(* IEC 61131-3 sources: deprecated-refusr-repo/samples (part 10) *)

(* ---- 4-MUX_towns-witty-ruing.st ---- *)
(*
This code implements a shuffled multiplexer with 4 control bits.
The control bits are: Data[N2], Data[N1], Data[N3], Data[N4]
The input bits are: Data[N7], Data[N5], Data[N6], Data[N12], Data[N15], Data[N10], Data[N8], Data[N13], Data[N18], Data[N9], Data[N11], Data[N14], Data[N17], Data[N19], Data[N16], Data[N20]

The symbolic expression is:
((((((((((((((((!((((!(IN2)) & (!(IN1))) & (!(IN3))) & (!(IN4)))) | IN7) & ((!(((IN2 & (!(IN1))) & (!(IN3))) & (!(IN4)))) | IN5)) & ((!((((!(IN2)) & IN1) & (!(IN3))) & (!(IN4)))) | IN6)) & ((!(((IN2 & IN1) & (!(IN3))) & (!(IN4)))) | IN12)) & ((!((((!(IN2)) & (!(IN1))) & IN3) & (!(IN4)))) | IN15)) & ((!(((IN2 & (!(IN1))) & IN3) & (!(IN4)))) | IN10)) & ((!((((!(IN2)) & IN1) & IN3) & (!(IN4)))) | IN8)) & ((!(((IN2 & IN1) & IN3) & (!(IN4)))) | IN13)) & ((!((((!(IN2)) & (!(IN1))) & (!(IN3))) & IN4)) | IN18)) & ((!(((IN2 & (!(IN1))) & (!(IN3))) & IN4)) | IN9)) & ((!((((!(IN2)) & IN1) & (!(IN3))) & IN4)) | IN11)) & ((!(((IN2 & IN1) & (!(IN3))) & IN4)) | IN14)) & ((!((((!(IN2)) & (!(IN1))) & IN3) & IN4)) | IN17)) & ((!(((IN2 & (!(IN1))) & IN3) & IN4)) | IN19)) & ((!((((!(IN2)) & IN1) & IN3) & IN4)) | IN16)) & ((!(((IN2 & IN1) & IN3) & IN4)) | IN20)

*)

FUNCTION_BLOCK F_CollectInput
  VAR_IN_OUT
      Data : ARRAY[1..20] OF BOOL;
  END_VAR
  VAR_INPUT
      TICK  : BOOL := 0;
      IN1   : BOOL := 0;
      IN2   : BOOL := 0;
      IN3   : BOOL := 0;
      IN4   : BOOL := 0;
      IN5   : BOOL := 0;
      RESET : BOOL := FALSE;
  END_VAR
  VAR_OUTPUT
      Finished : BOOL;
  END_VAR
  VAR
      j    : USINT := 1;
      tock : BOOL  := 0;
  END_VAR
  IF NOT RESET AND tock = NOT TICK THEN
      Data[j]   := IN1;
      Data[j+1] := IN2;
      Data[j+2] := IN3;
      Data[j+3] := IN4;
      Data[j+4] := IN5;
      j := j + 5;
      tock := TICK;
  ELSE
      j := 1;
      tock := 0;
  END_IF;
  Finished := (j > 20);
END_FUNCTION_BLOCK

PROGRAM Boiler
  VAR
    Data  : ARRAY[1..20] OF BOOL;
    Ready : BOOL;
    CollectInput : F_CollectInput;
  END_VAR
  VAR
    TICK     AT %IX1.0 : BOOL;
    IN1      AT %IX0.3 : BOOL;
    IN2      AT %IX0.4 : BOOL;
    IN3      AT %IX0.5 : BOOL;
    IN4      AT %IX0.6 : BOOL;
    IN5      AT %IX0.7 : BOOL;
    OutReady AT %QX0.0 : BOOL := FALSE;
    FeedNext AT %QX0.1 : BOOL := FALSE;
    Out      AT %QX0.2 : BOOL;
  END_VAR
  CollectInput(TICK:=TICK, IN1:=IN1, IN2:=IN2, IN3:=IN3, IN4:=IN4, IN5:=IN5);
  Ready := CollectInput.Finished;
  FeedNext := 1;
  IF Ready THEN
    Out := (((((((((((((((((NOT ((((NOT Data[2]) AND (NOT Data[1])) AND (NOT Data[3])) AND (NOT Data[4]))) OR Data[7]) AND ((NOT (((Data[2] AND (NOT Data[1])) AND (NOT Data[3])) AND (NOT Data[4]))) OR Data[5])) AND ((NOT ((((NOT Data[2]) AND Data[1]) AND (NOT Data[3])) AND (NOT Data[4]))) OR Data[6])) AND ((NOT (((Data[2] AND Data[1]) AND (NOT Data[3])) AND (NOT Data[4]))) OR Data[12])) AND ((NOT ((((NOT Data[2]) AND (NOT Data[1])) AND Data[3]) AND (NOT Data[4]))) OR Data[15])) AND ((NOT (((Data[2] AND (NOT Data[1])) AND Data[3]) AND (NOT Data[4]))) OR Data[10])) AND ((NOT ((((NOT Data[2]) AND Data[1]) AND Data[3]) AND (NOT Data[4]))) OR Data[8])) AND ((NOT (((Data[2] AND Data[1]) AND Data[3]) AND (NOT Data[4]))) OR Data[13])) AND ((NOT ((((NOT Data[2]) AND (NOT Data[1])) AND (NOT Data[3])) AND Data[4])) OR Data[18])) AND ((NOT (((Data[2] AND (NOT Data[1])) AND (NOT Data[3])) AND Data[4])) OR Data[9])) AND ((NOT ((((NOT Data[2]) AND Data[1]) AND (NOT Data[3])) AND Data[4])) OR Data[11])) AND ((NOT (((Data[2] AND Data[1]) AND (NOT Data[3])) AND Data[4])) OR Data[14])) AND ((NOT ((((NOT Data[2]) AND (NOT Data[1])) AND Data[3]) AND Data[4])) OR Data[17])) AND ((NOT (((Data[2] AND (NOT Data[1])) AND Data[3]) AND Data[4])) OR Data[19])) AND ((NOT ((((NOT Data[2]) AND Data[1]) AND Data[3]) AND Data[4])) OR Data[16])) AND ((NOT (((Data[2] AND Data[1]) AND Data[3]) AND Data[4])) OR Data[20]));
    OutReady := 1;
    CollectInput(RESET:=TRUE);
  END_IF;
END_PROGRAM

CONFIGURATION Config0
  RESOURCE Res0 ON PLC
    TASK task0(INTERVAL := T#20ms,PRIORITY := 0);
    PROGRAM instance0 WITH task0 : Boiler;
  END_RESOURCE
END_CONFIGURATION

(* ---- 4-MUX_tutti-shack-punky.st ---- *)
(*
This code implements a shuffled multiplexer with 4 control bits.
The control bits are: Data[N2], Data[N1], Data[N3], Data[N4]
The input bits are: Data[N5], Data[N6], Data[N9], Data[N7], Data[N11], Data[N8], Data[N10], Data[N12], Data[N13], Data[N14], Data[N16], Data[N17], Data[N15], Data[N18], Data[N19], Data[N20]

The symbolic expression is:
((((((((((((((((!((((!(IN2)) & (!(IN1))) & (!(IN3))) & (!(IN4)))) | IN5) & ((!(((IN2 & (!(IN1))) & (!(IN3))) & (!(IN4)))) | IN6)) & ((!((((!(IN2)) & IN1) & (!(IN3))) & (!(IN4)))) | IN9)) & ((!(((IN2 & IN1) & (!(IN3))) & (!(IN4)))) | IN7)) & ((!((((!(IN2)) & (!(IN1))) & IN3) & (!(IN4)))) | IN11)) & ((!(((IN2 & (!(IN1))) & IN3) & (!(IN4)))) | IN8)) & ((!((((!(IN2)) & IN1) & IN3) & (!(IN4)))) | IN10)) & ((!(((IN2 & IN1) & IN3) & (!(IN4)))) | IN12)) & ((!((((!(IN2)) & (!(IN1))) & (!(IN3))) & IN4)) | IN13)) & ((!(((IN2 & (!(IN1))) & (!(IN3))) & IN4)) | IN14)) & ((!((((!(IN2)) & IN1) & (!(IN3))) & IN4)) | IN16)) & ((!(((IN2 & IN1) & (!(IN3))) & IN4)) | IN17)) & ((!((((!(IN2)) & (!(IN1))) & IN3) & IN4)) | IN15)) & ((!(((IN2 & (!(IN1))) & IN3) & IN4)) | IN18)) & ((!((((!(IN2)) & IN1) & IN3) & IN4)) | IN19)) & ((!(((IN2 & IN1) & IN3) & IN4)) | IN20)

*)

FUNCTION_BLOCK F_CollectInput
  VAR_IN_OUT
      Data : ARRAY[1..20] OF BOOL;
  END_VAR
  VAR_INPUT
      TICK  : BOOL := 0;
      IN1   : BOOL := 0;
      IN2   : BOOL := 0;
      IN3   : BOOL := 0;
      IN4   : BOOL := 0;
      IN5   : BOOL := 0;
      RESET : BOOL := FALSE;
  END_VAR
  VAR_OUTPUT
      Finished : BOOL;
  END_VAR
  VAR
      j    : USINT := 1;
      tock : BOOL  := 0;
  END_VAR
  IF NOT RESET AND tock = NOT TICK THEN
      Data[j]   := IN1;
      Data[j+1] := IN2;
      Data[j+2] := IN3;
      Data[j+3] := IN4;
      Data[j+4] := IN5;
      j := j + 5;
      tock := TICK;
  ELSE
      j := 1;
      tock := 0;
  END_IF;
  Finished := (j > 20);
END_FUNCTION_BLOCK

PROGRAM Boiler
  VAR
    Data  : ARRAY[1..20] OF BOOL;
    Ready : BOOL;
    CollectInput : F_CollectInput;
  END_VAR
  VAR
    TICK     AT %IX1.0 : BOOL;
    IN1      AT %IX0.3 : BOOL;
    IN2      AT %IX0.4 : BOOL;
    IN3      AT %IX0.5 : BOOL;
    IN4      AT %IX0.6 : BOOL;
    IN5      AT %IX0.7 : BOOL;
    OutReady AT %QX0.0 : BOOL := FALSE;
    FeedNext AT %QX0.1 : BOOL := FALSE;
    Out      AT %QX0.2 : BOOL;
  END_VAR
  CollectInput(TICK:=TICK, IN1:=IN1, IN2:=IN2, IN3:=IN3, IN4:=IN4, IN5:=IN5);
  Ready := CollectInput.Finished;
  FeedNext := 1;
  IF Ready THEN
    Out := (((((((((((((((((NOT ((((NOT Data[2]) AND (NOT Data[1])) AND (NOT Data[3])) AND (NOT Data[4]))) OR Data[5]) AND ((NOT (((Data[2] AND (NOT Data[1])) AND (NOT Data[3])) AND (NOT Data[4]))) OR Data[6])) AND ((NOT ((((NOT Data[2]) AND Data[1]) AND (NOT Data[3])) AND (NOT Data[4]))) OR Data[9])) AND ((NOT (((Data[2] AND Data[1]) AND (NOT Data[3])) AND (NOT Data[4]))) OR Data[7])) AND ((NOT ((((NOT Data[2]) AND (NOT Data[1])) AND Data[3]) AND (NOT Data[4]))) OR Data[11])) AND ((NOT (((Data[2] AND (NOT Data[1])) AND Data[3]) AND (NOT Data[4]))) OR Data[8])) AND ((NOT ((((NOT Data[2]) AND Data[1]) AND Data[3]) AND (NOT Data[4]))) OR Data[10])) AND ((NOT (((Data[2] AND Data[1]) AND Data[3]) AND (NOT Data[4]))) OR Data[12])) AND ((NOT ((((NOT Data[2]) AND (NOT Data[1])) AND (NOT Data[3])) AND Data[4])) OR Data[13])) AND ((NOT (((Data[2] AND (NOT Data[1])) AND (NOT Data[3])) AND Data[4])) OR Data[14])) AND ((NOT ((((NOT Data[2]) AND Data[1]) AND (NOT Data[3])) AND Data[4])) OR Data[16])) AND ((NOT (((Data[2] AND Data[1]) AND (NOT Data[3])) AND Data[4])) OR Data[17])) AND ((NOT ((((NOT Data[2]) AND (NOT Data[1])) AND Data[3]) AND Data[4])) OR Data[15])) AND ((NOT (((Data[2] AND (NOT Data[1])) AND Data[3]) AND Data[4])) OR Data[18])) AND ((NOT ((((NOT Data[2]) AND Data[1]) AND Data[3]) AND Data[4])) OR Data[19])) AND ((NOT (((Data[2] AND Data[1]) AND Data[3]) AND Data[4])) OR Data[20]));
    OutReady := 1;
    CollectInput(RESET:=TRUE);
  END_IF;
END_PROGRAM

CONFIGURATION Config0
  RESOURCE Res0 ON PLC
    TASK task0(INTERVAL := T#20ms,PRIORITY := 0);
    PROGRAM instance0 WITH task0 : Boiler;
  END_RESOURCE
END_CONFIGURATION

(* ---- 4-MUX_tweed-dweeb-warns.st ---- *)
(*
This code implements a shuffled multiplexer with 4 control bits.
The control bits are: Data[N5], Data[N1], Data[N2], Data[N3]
The input bits are: Data[N4], Data[N6], Data[N8], Data[N9], Data[N7], Data[N11], Data[N13], Data[N10], Data[N12], Data[N14], Data[N17], Data[N15], Data[N16], Data[N19], Data[N20], Data[N18]

The symbolic expression is:
((((((((((((((((!((((!(IN5)) & (!(IN1))) & (!(IN2))) & (!(IN3)))) | IN4) & ((!(((IN5 & (!(IN1))) & (!(IN2))) & (!(IN3)))) | IN6)) & ((!((((!(IN5)) & IN1) & (!(IN2))) & (!(IN3)))) | IN8)) & ((!(((IN5 & IN1) & (!(IN2))) & (!(IN3)))) | IN9)) & ((!((((!(IN5)) & (!(IN1))) & IN2) & (!(IN3)))) | IN7)) & ((!(((IN5 & (!(IN1))) & IN2) & (!(IN3)))) | IN11)) & ((!((((!(IN5)) & IN1) & IN2) & (!(IN3)))) | IN13)) & ((!(((IN5 & IN1) & IN2) & (!(IN3)))) | IN10)) & ((!((((!(IN5)) & (!(IN1))) & (!(IN2))) & IN3)) | IN12)) & ((!(((IN5 & (!(IN1))) & (!(IN2))) & IN3)) | IN14)) & ((!((((!(IN5)) & IN1) & (!(IN2))) & IN3)) | IN17)) & ((!(((IN5 & IN1) & (!(IN2))) & IN3)) | IN15)) & ((!((((!(IN5)) & (!(IN1))) & IN2) & IN3)) | IN16)) & ((!(((IN5 & (!(IN1))) & IN2) & IN3)) | IN19)) & ((!((((!(IN5)) & IN1) & IN2) & IN3)) | IN20)) & ((!(((IN5 & IN1) & IN2) & IN3)) | IN18)

*)

FUNCTION_BLOCK F_CollectInput
  VAR_IN_OUT
      Data : ARRAY[1..20] OF BOOL;
  END_VAR
  VAR_INPUT
      TICK  : BOOL := 0;
      IN1   : BOOL := 0;
      IN2   : BOOL := 0;
      IN3   : BOOL := 0;
      IN4   : BOOL := 0;
      IN5   : BOOL := 0;
      RESET : BOOL := FALSE;
  END_VAR
  VAR_OUTPUT
      Finished : BOOL;
  END_VAR
  VAR
      j    : USINT := 1;
      tock : BOOL  := 0;
  END_VAR
  IF NOT RESET AND tock = NOT TICK THEN
      Data[j]   := IN1;
      Data[j+1] := IN2;
      Data[j+2] := IN3;
      Data[j+3] := IN4;
      Data[j+4] := IN5;
      j := j + 5;
      tock := TICK;
  ELSE
      j := 1;
      tock := 0;
  END_IF;
  Finished := (j > 20);
END_FUNCTION_BLOCK

PROGRAM Boiler
  VAR
    Data  : ARRAY[1..20] OF BOOL;
    Ready : BOOL;
    CollectInput : F_CollectInput;
  END_VAR
  VAR
    TICK     AT %IX1.0 : BOOL;
    IN1      AT %IX0.3 : BOOL;
    IN2      AT %IX0.4 : BOOL;
    IN3      AT %IX0.5 : BOOL;
    IN4      AT %IX0.6 : BOOL;
    IN5      AT %IX0.7 : BOOL;
    OutReady AT %QX0.0 : BOOL := FALSE;
    FeedNext AT %QX0.1 : BOOL := FALSE;
    Out      AT %QX0.2 : BOOL;
  END_VAR
  CollectInput(TICK:=TICK, IN1:=IN1, IN2:=IN2, IN3:=IN3, IN4:=IN4, IN5:=IN5);
  Ready := CollectInput.Finished;
  FeedNext := 1;
  IF Ready THEN
    Out := (((((((((((((((((NOT ((((NOT Data[5]) AND (NOT Data[1])) AND (NOT Data[2])) AND (NOT Data[3]))) OR Data[4]) AND ((NOT (((Data[5] AND (NOT Data[1])) AND (NOT Data[2])) AND (NOT Data[3]))) OR Data[6])) AND ((NOT ((((NOT Data[5]) AND Data[1]) AND (NOT Data[2])) AND (NOT Data[3]))) OR Data[8])) AND ((NOT (((Data[5] AND Data[1]) AND (NOT Data[2])) AND (NOT Data[3]))) OR Data[9])) AND ((NOT ((((NOT Data[5]) AND (NOT Data[1])) AND Data[2]) AND (NOT Data[3]))) OR Data[7])) AND ((NOT (((Data[5] AND (NOT Data[1])) AND Data[2]) AND (NOT Data[3]))) OR Data[11])) AND ((NOT ((((NOT Data[5]) AND Data[1]) AND Data[2]) AND (NOT Data[3]))) OR Data[13])) AND ((NOT (((Data[5] AND Data[1]) AND Data[2]) AND (NOT Data[3]))) OR Data[10])) AND ((NOT ((((NOT Data[5]) AND (NOT Data[1])) AND (NOT Data[2])) AND Data[3])) OR Data[12])) AND ((NOT (((Data[5] AND (NOT Data[1])) AND (NOT Data[2])) AND Data[3])) OR Data[14])) AND ((NOT ((((NOT Data[5]) AND Data[1]) AND (NOT Data[2])) AND Data[3])) OR Data[17])) AND ((NOT (((Data[5] AND Data[1]) AND (NOT Data[2])) AND Data[3])) OR Data[15])) AND ((NOT ((((NOT Data[5]) AND (NOT Data[1])) AND Data[2]) AND Data[3])) OR Data[16])) AND ((NOT (((Data[5] AND (NOT Data[1])) AND Data[2]) AND Data[3])) OR Data[19])) AND ((NOT ((((NOT Data[5]) AND Data[1]) AND Data[2]) AND Data[3])) OR Data[20])) AND ((NOT (((Data[5] AND Data[1]) AND Data[2]) AND Data[3])) OR Data[18]));
    OutReady := 1;
    CollectInput(RESET:=TRUE);
  END_IF;
END_PROGRAM

CONFIGURATION Config0
  RESOURCE Res0 ON PLC
    TASK task0(INTERVAL := T#20ms,PRIORITY := 0);
    PROGRAM instance0 WITH task0 : Boiler;
  END_RESOURCE
END_CONFIGURATION

(* ---- 4-MUX_tweed-nitty-duels.st ---- *)
(*
This code implements a shuffled multiplexer with 4 control bits.
The control bits are: Data[N1], Data[N2], Data[N9], Data[N3]
The input bits are: Data[N5], Data[N4], Data[N8], Data[N7], Data[N6], Data[N17], Data[N14], Data[N18], Data[N10], Data[N11], Data[N12], Data[N13], Data[N19], Data[N15], Data[N20], Data[N16]

The symbolic expression is:
((((((((((((((((!((((!(IN1)) & (!(IN2))) & (!(IN9))) & (!(IN3)))) | IN5) & ((!(((IN1 & (!(IN2))) & (!(IN9))) & (!(IN3)))) | IN4)) & ((!((((!(IN1)) & IN2) & (!(IN9))) & (!(IN3)))) | IN8)) & ((!(((IN1 & IN2) & (!(IN9))) & (!(IN3)))) | IN7)) & ((!((((!(IN1)) & (!(IN2))) & IN9) & (!(IN3)))) | IN6)) & ((!(((IN1 & (!(IN2))) & IN9) & (!(IN3)))) | IN17)) & ((!((((!(IN1)) & IN2) & IN9) & (!(IN3)))) | IN14)) & ((!(((IN1 & IN2) & IN9) & (!(IN3)))) | IN18)) & ((!((((!(IN1)) & (!(IN2))) & (!(IN9))) & IN3)) | IN10)) & ((!(((IN1 & (!(IN2))) & (!(IN9))) & IN3)) | IN11)) & ((!((((!(IN1)) & IN2) & (!(IN9))) & IN3)) | IN12)) & ((!(((IN1 & IN2) & (!(IN9))) & IN3)) | IN13)) & ((!((((!(IN1)) & (!(IN2))) & IN9) & IN3)) | IN19)) & ((!(((IN1 & (!(IN2))) & IN9) & IN3)) | IN15)) & ((!((((!(IN1)) & IN2) & IN9) & IN3)) | IN20)) & ((!(((IN1 & IN2) & IN9) & IN3)) | IN16)

*)

FUNCTION_BLOCK F_CollectInput
  VAR_IN_OUT
      Data : ARRAY[1..20] OF BOOL;
  END_VAR
  VAR_INPUT
      TICK  : BOOL := 0;
      IN1   : BOOL := 0;
      IN2   : BOOL := 0;
      IN3   : BOOL := 0;
      IN4   : BOOL := 0;
      IN5   : BOOL := 0;
      RESET : BOOL := FALSE;
  END_VAR
  VAR_OUTPUT
      Finished : BOOL;
  END_VAR
  VAR
      j    : USINT := 1;
      tock : BOOL  := 0;
  END_VAR
  IF NOT RESET AND tock = NOT TICK THEN
      Data[j]   := IN1;
      Data[j+1] := IN2;
      Data[j+2] := IN3;
      Data[j+3] := IN4;
      Data[j+4] := IN5;
      j := j + 5;
      tock := TICK;
  ELSE
      j := 1;
      tock := 0;
  END_IF;
  Finished := (j > 20);
END_FUNCTION_BLOCK

PROGRAM Boiler
  VAR
    Data  : ARRAY[1..20] OF BOOL;
    Ready : BOOL;
    CollectInput : F_CollectInput;
  END_VAR
  VAR
    TICK     AT %IX1.0 : BOOL;
    IN1      AT %IX0.3 : BOOL;
    IN2      AT %IX0.4 : BOOL;
    IN3      AT %IX0.5 : BOOL;
    IN4      AT %IX0.6 : BOOL;
    IN5      AT %IX0.7 : BOOL;
    OutReady AT %QX0.0 : BOOL := FALSE;
    FeedNext AT %QX0.1 : BOOL := FALSE;
    Out      AT %QX0.2 : BOOL;
  END_VAR
  CollectInput(TICK:=TICK, IN1:=IN1, IN2:=IN2, IN3:=IN3, IN4:=IN4, IN5:=IN5);
  Ready := CollectInput.Finished;
  FeedNext := 1;
  IF Ready THEN
    Out := (((((((((((((((((NOT ((((NOT Data[1]) AND (NOT Data[2])) AND (NOT Data[9])) AND (NOT Data[3]))) OR Data[5]) AND ((NOT (((Data[1] AND (NOT Data[2])) AND (NOT Data[9])) AND (NOT Data[3]))) OR Data[4])) AND ((NOT ((((NOT Data[1]) AND Data[2]) AND (NOT Data[9])) AND (NOT Data[3]))) OR Data[8])) AND ((NOT (((Data[1] AND Data[2]) AND (NOT Data[9])) AND (NOT Data[3]))) OR Data[7])) AND ((NOT ((((NOT Data[1]) AND (NOT Data[2])) AND Data[9]) AND (NOT Data[3]))) OR Data[6])) AND ((NOT (((Data[1] AND (NOT Data[2])) AND Data[9]) AND (NOT Data[3]))) OR Data[17])) AND ((NOT ((((NOT Data[1]) AND Data[2]) AND Data[9]) AND (NOT Data[3]))) OR Data[14])) AND ((NOT (((Data[1] AND Data[2]) AND Data[9]) AND (NOT Data[3]))) OR Data[18])) AND ((NOT ((((NOT Data[1]) AND (NOT Data[2])) AND (NOT Data[9])) AND Data[3])) OR Data[10])) AND ((NOT (((Data[1] AND (NOT Data[2])) AND (NOT Data[9])) AND Data[3])) OR Data[11])) AND ((NOT ((((NOT Data[1]) AND Data[2]) AND (NOT Data[9])) AND Data[3])) OR Data[12])) AND ((NOT (((Data[1] AND Data[2]) AND (NOT Data[9])) AND Data[3])) OR Data[13])) AND ((NOT ((((NOT Data[1]) AND (NOT Data[2])) AND Data[9]) AND Data[3])) OR Data[19])) AND ((NOT (((Data[1] AND (NOT Data[2])) AND Data[9]) AND Data[3])) OR Data[15])) AND ((NOT ((((NOT Data[1]) AND Data[2]) AND Data[9]) AND Data[3])) OR Data[20])) AND ((NOT (((Data[1] AND Data[2]) AND Data[9]) AND Data[3])) OR Data[16]));
    OutReady := 1;
    CollectInput(RESET:=TRUE);
  END_IF;
END_PROGRAM

CONFIGURATION Config0
  RESOURCE Res0 ON PLC
    TASK task0(INTERVAL := T#20ms,PRIORITY := 0);
    PROGRAM instance0 WITH task0 : Boiler;
  END_RESOURCE
END_CONFIGURATION

(* ---- 4-MUX_twice-mined-dimes.st ---- *)
(*
This code implements a shuffled multiplexer with 4 control bits.
The control bits are: Data[N1], Data[N2], Data[N3], Data[N5]
The input bits are: Data[N9], Data[N4], Data[N14], Data[N6], Data[N7], Data[N8], Data[N10], Data[N11], Data[N15], Data[N12], Data[N13], Data[N16], Data[N19], Data[N17], Data[N20], Data[N18]

The symbolic expression is:
((((((((((((((((!((((!(IN1)) & (!(IN2))) & (!(IN3))) & (!(IN5)))) | IN9) & ((!(((IN1 & (!(IN2))) & (!(IN3))) & (!(IN5)))) | IN4)) & ((!((((!(IN1)) & IN2) & (!(IN3))) & (!(IN5)))) | IN14)) & ((!(((IN1 & IN2) & (!(IN3))) & (!(IN5)))) | IN6)) & ((!((((!(IN1)) & (!(IN2))) & IN3) & (!(IN5)))) | IN7)) & ((!(((IN1 & (!(IN2))) & IN3) & (!(IN5)))) | IN8)) & ((!((((!(IN1)) & IN2) & IN3) & (!(IN5)))) | IN10)) & ((!(((IN1 & IN2) & IN3) & (!(IN5)))) | IN11)) & ((!((((!(IN1)) & (!(IN2))) & (!(IN3))) & IN5)) | IN15)) & ((!(((IN1 & (!(IN2))) & (!(IN3))) & IN5)) | IN12)) & ((!((((!(IN1)) & IN2) & (!(IN3))) & IN5)) | IN13)) & ((!(((IN1 & IN2) & (!(IN3))) & IN5)) | IN16)) & ((!((((!(IN1)) & (!(IN2))) & IN3) & IN5)) | IN19)) & ((!(((IN1 & (!(IN2))) & IN3) & IN5)) | IN17)) & ((!((((!(IN1)) & IN2) & IN3) & IN5)) | IN20)) & ((!(((IN1 & IN2) & IN3) & IN5)) | IN18)

*)

FUNCTION_BLOCK F_CollectInput
  VAR_IN_OUT
      Data : ARRAY[1..20] OF BOOL;
  END_VAR
  VAR_INPUT
      TICK  : BOOL := 0;
      IN1   : BOOL := 0;
      IN2   : BOOL := 0;
      IN3   : BOOL := 0;
      IN4   : BOOL := 0;
      IN5   : BOOL := 0;
      RESET : BOOL := FALSE;
  END_VAR
  VAR_OUTPUT
      Finished : BOOL;
  END_VAR
  VAR
      j    : USINT := 1;
      tock : BOOL  := 0;
  END_VAR
  IF NOT RESET AND tock = NOT TICK THEN
      Data[j]   := IN1;
      Data[j+1] := IN2;
      Data[j+2] := IN3;
      Data[j+3] := IN4;
      Data[j+4] := IN5;
      j := j + 5;
      tock := TICK;
  ELSE
      j := 1;
      tock := 0;
  END_IF;
  Finished := (j > 20);
END_FUNCTION_BLOCK

PROGRAM Boiler
  VAR
    Data  : ARRAY[1..20] OF BOOL;
    Ready : BOOL;
    CollectInput : F_CollectInput;
  END_VAR
  VAR
    TICK     AT %IX1.0 : BOOL;
    IN1      AT %IX0.3 : BOOL;
    IN2      AT %IX0.4 : BOOL;
    IN3      AT %IX0.5 : BOOL;
    IN4      AT %IX0.6 : BOOL;
    IN5      AT %IX0.7 : BOOL;
    OutReady AT %QX0.0 : BOOL := FALSE;
    FeedNext AT %QX0.1 : BOOL := FALSE;
    Out      AT %QX0.2 : BOOL;
  END_VAR
  CollectInput(TICK:=TICK, IN1:=IN1, IN2:=IN2, IN3:=IN3, IN4:=IN4, IN5:=IN5);
  Ready := CollectInput.Finished;
  FeedNext := 1;
  IF Ready THEN
    Out := (((((((((((((((((NOT ((((NOT Data[1]) AND (NOT Data[2])) AND (NOT Data[3])) AND (NOT Data[5]))) OR Data[9]) AND ((NOT (((Data[1] AND (NOT Data[2])) AND (NOT Data[3])) AND (NOT Data[5]))) OR Data[4])) AND ((NOT ((((NOT Data[1]) AND Data[2]) AND (NOT Data[3])) AND (NOT Data[5]))) OR Data[14])) AND ((NOT (((Data[1] AND Data[2]) AND (NOT Data[3])) AND (NOT Data[5]))) OR Data[6])) AND ((NOT ((((NOT Data[1]) AND (NOT Data[2])) AND Data[3]) AND (NOT Data[5]))) OR Data[7])) AND ((NOT (((Data[1] AND (NOT Data[2])) AND Data[3]) AND (NOT Data[5]))) OR Data[8])) AND ((NOT ((((NOT Data[1]) AND Data[2]) AND Data[3]) AND (NOT Data[5]))) OR Data[10])) AND ((NOT (((Data[1] AND Data[2]) AND Data[3]) AND (NOT Data[5]))) OR Data[11])) AND ((NOT ((((NOT Data[1]) AND (NOT Data[2])) AND (NOT Data[3])) AND Data[5])) OR Data[15])) AND ((NOT (((Data[1] AND (NOT Data[2])) AND (NOT Data[3])) AND Data[5])) OR Data[12])) AND ((NOT ((((NOT Data[1]) AND Data[2]) AND (NOT Data[3])) AND Data[5])) OR Data[13])) AND ((NOT (((Data[1] AND Data[2]) AND (NOT Data[3])) AND Data[5])) OR Data[16])) AND ((NOT ((((NOT Data[1]) AND (NOT Data[2])) AND Data[3]) AND Data[5])) OR Data[19])) AND ((NOT (((Data[1] AND (NOT Data[2])) AND Data[3]) AND Data[5])) OR Data[17])) AND ((NOT ((((NOT Data[1]) AND Data[2]) AND Data[3]) AND Data[5])) OR Data[20])) AND ((NOT (((Data[1] AND Data[2]) AND Data[3]) AND Data[5])) OR Data[18]));
    OutReady := 1;
    CollectInput(RESET:=TRUE);
  END_IF;
END_PROGRAM

CONFIGURATION Config0
  RESOURCE Res0 ON PLC
    TASK task0(INTERVAL := T#20ms,PRIORITY := 0);
    PROGRAM instance0 WITH task0 : Boiler;
  END_RESOURCE
END_CONFIGURATION

(* ---- 4-MUX_twine-odder-crimp.st ---- *)
(*
This code implements a shuffled multiplexer with 4 control bits.
The control bits are: Data[N2], Data[N4], Data[N3], Data[N5]
The input bits are: Data[N1], Data[N11], Data[N6], Data[N7], Data[N8], Data[N9], Data[N12], Data[N17], Data[N14], Data[N18], Data[N10], Data[N13], Data[N15], Data[N16], Data[N19], Data[N20]

The symbolic expression is:
((((((((((((((((!((((!(IN2)) & (!(IN4))) & (!(IN3))) & (!(IN5)))) | IN1) & ((!(((IN2 & (!(IN4))) & (!(IN3))) & (!(IN5)))) | IN11)) & ((!((((!(IN2)) & IN4) & (!(IN3))) & (!(IN5)))) | IN6)) & ((!(((IN2 & IN4) & (!(IN3))) & (!(IN5)))) | IN7)) & ((!((((!(IN2)) & (!(IN4))) & IN3) & (!(IN5)))) | IN8)) & ((!(((IN2 & (!(IN4))) & IN3) & (!(IN5)))) | IN9)) & ((!((((!(IN2)) & IN4) & IN3) & (!(IN5)))) | IN12)) & ((!(((IN2 & IN4) & IN3) & (!(IN5)))) | IN17)) & ((!((((!(IN2)) & (!(IN4))) & (!(IN3))) & IN5)) | IN14)) & ((!(((IN2 & (!(IN4))) & (!(IN3))) & IN5)) | IN18)) & ((!((((!(IN2)) & IN4) & (!(IN3))) & IN5)) | IN10)) & ((!(((IN2 & IN4) & (!(IN3))) & IN5)) | IN13)) & ((!((((!(IN2)) & (!(IN4))) & IN3) & IN5)) | IN15)) & ((!(((IN2 & (!(IN4))) & IN3) & IN5)) | IN16)) & ((!((((!(IN2)) & IN4) & IN3) & IN5)) | IN19)) & ((!(((IN2 & IN4) & IN3) & IN5)) | IN20)

*)

FUNCTION_BLOCK F_CollectInput
  VAR_IN_OUT
      Data : ARRAY[1..20] OF BOOL;
  END_VAR
  VAR_INPUT
      TICK  : BOOL := 0;
      IN1   : BOOL := 0;
      IN2   : BOOL := 0;
      IN3   : BOOL := 0;
      IN4   : BOOL := 0;
      IN5   : BOOL := 0;
      RESET : BOOL := FALSE;
  END_VAR
  VAR_OUTPUT
      Finished : BOOL;
  END_VAR
  VAR
      j    : USINT := 1;
      tock : BOOL  := 0;
  END_VAR
  IF NOT RESET AND tock = NOT TICK THEN
      Data[j]   := IN1;
      Data[j+1] := IN2;
      Data[j+2] := IN3;
      Data[j+3] := IN4;
      Data[j+4] := IN5;
      j := j + 5;
      tock := TICK;
  ELSE
      j := 1;
      tock := 0;
  END_IF;
  Finished := (j > 20);
END_FUNCTION_BLOCK

PROGRAM Boiler
  VAR
    Data  : ARRAY[1..20] OF BOOL;
    Ready : BOOL;
    CollectInput : F_CollectInput;
  END_VAR
  VAR
    TICK     AT %IX1.0 : BOOL;
    IN1      AT %IX0.3 : BOOL;
    IN2      AT %IX0.4 : BOOL;
    IN3      AT %IX0.5 : BOOL;
    IN4      AT %IX0.6 : BOOL;
    IN5      AT %IX0.7 : BOOL;
    OutReady AT %QX0.0 : BOOL := FALSE;
    FeedNext AT %QX0.1 : BOOL := FALSE;
    Out      AT %QX0.2 : BOOL;
  END_VAR
  CollectInput(TICK:=TICK, IN1:=IN1, IN2:=IN2, IN3:=IN3, IN4:=IN4, IN5:=IN5);
  Ready := CollectInput.Finished;
  FeedNext := 1;
  IF Ready THEN
    Out := (((((((((((((((((NOT ((((NOT Data[2]) AND (NOT Data[4])) AND (NOT Data[3])) AND (NOT Data[5]))) OR Data[1]) AND ((NOT (((Data[2] AND (NOT Data[4])) AND (NOT Data[3])) AND (NOT Data[5]))) OR Data[11])) AND ((NOT ((((NOT Data[2]) AND Data[4]) AND (NOT Data[3])) AND (NOT Data[5]))) OR Data[6])) AND ((NOT (((Data[2] AND Data[4]) AND (NOT Data[3])) AND (NOT Data[5]))) OR Data[7])) AND ((NOT ((((NOT Data[2]) AND (NOT Data[4])) AND Data[3]) AND (NOT Data[5]))) OR Data[8])) AND ((NOT (((Data[2] AND (NOT Data[4])) AND Data[3]) AND (NOT Data[5]))) OR Data[9])) AND ((NOT ((((NOT Data[2]) AND Data[4]) AND Data[3]) AND (NOT Data[5]))) OR Data[12])) AND ((NOT (((Data[2] AND Data[4]) AND Data[3]) AND (NOT Data[5]))) OR Data[17])) AND ((NOT ((((NOT Data[2]) AND (NOT Data[4])) AND (NOT Data[3])) AND Data[5])) OR Data[14])) AND ((NOT (((Data[2] AND (NOT Data[4])) AND (NOT Data[3])) AND Data[5])) OR Data[18])) AND ((NOT ((((NOT Data[2]) AND Data[4]) AND (NOT Data[3])) AND Data[5])) OR Data[10])) AND ((NOT (((Data[2] AND Data[4]) AND (NOT Data[3])) AND Data[5])) OR Data[13])) AND ((NOT ((((NOT Data[2]) AND (NOT Data[4])) AND Data[3]) AND Data[5])) OR Data[15])) AND ((NOT (((Data[2] AND (NOT Data[4])) AND Data[3]) AND Data[5])) OR Data[16])) AND ((NOT ((((NOT Data[2]) AND Data[4]) AND Data[3]) AND Data[5])) OR Data[19])) AND ((NOT (((Data[2] AND Data[4]) AND Data[3]) AND Data[5])) OR Data[20]));
    OutReady := 1;
    CollectInput(RESET:=TRUE);
  END_IF;
END_PROGRAM

CONFIGURATION Config0
  RESOURCE Res0 ON PLC
    TASK task0(INTERVAL := T#20ms,PRIORITY := 0);
    PROGRAM instance0 WITH task0 : Boiler;
  END_RESOURCE
END_CONFIGURATION

(* ---- 4-MUX_warty-auric-paren.st ---- *)
(*
This code implements a shuffled multiplexer with 4 control bits.
The control bits are: Data[N2], Data[N1], Data[N11], Data[N3]
The input bits are: Data[N4], Data[N5], Data[N7], Data[N12], Data[N8], Data[N10], Data[N6], Data[N9], Data[N14], Data[N16], Data[N18], Data[N15], Data[N17], Data[N19], Data[N20], Data[N13]

The symbolic expression is:
((((((((((((((((!((((!(IN2)) & (!(IN1))) & (!(IN11))) & (!(IN3)))) | IN4) & ((!(((IN2 & (!(IN1))) & (!(IN11))) & (!(IN3)))) | IN5)) & ((!((((!(IN2)) & IN1) & (!(IN11))) & (!(IN3)))) | IN7)) & ((!(((IN2 & IN1) & (!(IN11))) & (!(IN3)))) | IN12)) & ((!((((!(IN2)) & (!(IN1))) & IN11) & (!(IN3)))) | IN8)) & ((!(((IN2 & (!(IN1))) & IN11) & (!(IN3)))) | IN10)) & ((!((((!(IN2)) & IN1) & IN11) & (!(IN3)))) | IN6)) & ((!(((IN2 & IN1) & IN11) & (!(IN3)))) | IN9)) & ((!((((!(IN2)) & (!(IN1))) & (!(IN11))) & IN3)) | IN14)) & ((!(((IN2 & (!(IN1))) & (!(IN11))) & IN3)) | IN16)) & ((!((((!(IN2)) & IN1) & (!(IN11))) & IN3)) | IN18)) & ((!(((IN2 & IN1) & (!(IN11))) & IN3)) | IN15)) & ((!((((!(IN2)) & (!(IN1))) & IN11) & IN3)) | IN17)) & ((!(((IN2 & (!(IN1))) & IN11) & IN3)) | IN19)) & ((!((((!(IN2)) & IN1) & IN11) & IN3)) | IN20)) & ((!(((IN2 & IN1) & IN11) & IN3)) | IN13)

*)

FUNCTION_BLOCK F_CollectInput
  VAR_IN_OUT
      Data : ARRAY[1..20] OF BOOL;
  END_VAR
  VAR_INPUT
      TICK  : BOOL := 0;
      IN1   : BOOL := 0;
      IN2   : BOOL := 0;
      IN3   : BOOL := 0;
      IN4   : BOOL := 0;
      IN5   : BOOL := 0;
      RESET : BOOL := FALSE;
  END_VAR
  VAR_OUTPUT
      Finished : BOOL;
  END_VAR
  VAR
      j    : USINT := 1;
      tock : BOOL  := 0;
  END_VAR
  IF NOT RESET AND tock = NOT TICK THEN
      Data[j]   := IN1;
      Data[j+1] := IN2;
      Data[j+2] := IN3;
      Data[j+3] := IN4;
      Data[j+4] := IN5;
      j := j + 5;
      tock := TICK;
  ELSE
      j := 1;
      tock := 0;
  END_IF;
  Finished := (j > 20);
END_FUNCTION_BLOCK

PROGRAM Boiler
  VAR
    Data  : ARRAY[1..20] OF BOOL;
    Ready : BOOL;
    CollectInput : F_CollectInput;
  END_VAR
  VAR
    TICK     AT %IX1.0 : BOOL;
    IN1      AT %IX0.3 : BOOL;
    IN2      AT %IX0.4 : BOOL;
    IN3      AT %IX0.5 : BOOL;
    IN4      AT %IX0.6 : BOOL;
    IN5      AT %IX0.7 : BOOL;
    OutReady AT %QX0.0 : BOOL := FALSE;
    FeedNext AT %QX0.1 : BOOL := FALSE;
    Out      AT %QX0.2 : BOOL;
  END_VAR
  CollectInput(TICK:=TICK, IN1:=IN1, IN2:=IN2, IN3:=IN3, IN4:=IN4, IN5:=IN5);
  Ready := CollectInput.Finished;
  FeedNext := 1;
  IF Ready THEN
    Out := (((((((((((((((((NOT ((((NOT Data[2]) AND (NOT Data[1])) AND (NOT Data[11])) AND (NOT Data[3]))) OR Data[4]) AND ((NOT (((Data[2] AND (NOT Data[1])) AND (NOT Data[11])) AND (NOT Data[3]))) OR Data[5])) AND ((NOT ((((NOT Data[2]) AND Data[1]) AND (NOT Data[11])) AND (NOT Data[3]))) OR Data[7])) AND ((NOT (((Data[2] AND Data[1]) AND (NOT Data[11])) AND (NOT Data[3]))) OR Data[12])) AND ((NOT ((((NOT Data[2]) AND (NOT Data[1])) AND Data[11]) AND (NOT Data[3]))) OR Data[8])) AND ((NOT (((Data[2] AND (NOT Data[1])) AND Data[11]) AND (NOT Data[3]))) OR Data[10])) AND ((NOT ((((NOT Data[2]) AND Data[1]) AND Data[11]) AND (NOT Data[3]))) OR Data[6])) AND ((NOT (((Data[2] AND Data[1]) AND Data[11]) AND (NOT Data[3]))) OR Data[9])) AND ((NOT ((((NOT Data[2]) AND (NOT Data[1])) AND (NOT Data[11])) AND Data[3])) OR Data[14])) AND ((NOT (((Data[2] AND (NOT Data[1])) AND (NOT Data[11])) AND Data[3])) OR Data[16])) AND ((NOT ((((NOT Data[2]) AND Data[1]) AND (NOT Data[11])) AND Data[3])) OR Data[18])) AND ((NOT (((Data[2] AND Data[1]) AND (NOT Data[11])) AND Data[3])) OR Data[15])) AND ((NOT ((((NOT Data[2]) AND (NOT Data[1])) AND Data[11]) AND Data[3])) OR Data[17])) AND ((NOT (((Data[2] AND (NOT Data[1])) AND Data[11]) AND Data[3])) OR Data[19])) AND ((NOT ((((NOT Data[2]) AND Data[1]) AND Data[11]) AND Data[3])) OR Data[20])) AND ((NOT (((Data[2] AND Data[1]) AND Data[11]) AND Data[3])) OR Data[13]));
    OutReady := 1;
    CollectInput(RESET:=TRUE);
  END_IF;
END_PROGRAM

CONFIGURATION Config0
  RESOURCE Res0 ON PLC
    TASK task0(INTERVAL := T#20ms,PRIORITY := 0);
    PROGRAM instance0 WITH task0 : Boiler;
  END_RESOURCE
END_CONFIGURATION

(* ---- 4-MUX_weest-tombs-frosh.st ---- *)
(*
This code implements a shuffled multiplexer with 4 control bits.
The control bits are: Data[N2], Data[N1], Data[N3], Data[N5]
The input bits are: Data[N6], Data[N7], Data[N9], Data[N8], Data[N11], Data[N4], Data[N13], Data[N10], Data[N12], Data[N18], Data[N16], Data[N14], Data[N15], Data[N17], Data[N19], Data[N20]

The symbolic expression is:
((((((((((((((((!((((!(IN2)) & (!(IN1))) & (!(IN3))) & (!(IN5)))) | IN6) & ((!(((IN2 & (!(IN1))) & (!(IN3))) & (!(IN5)))) | IN7)) & ((!((((!(IN2)) & IN1) & (!(IN3))) & (!(IN5)))) | IN9)) & ((!(((IN2 & IN1) & (!(IN3))) & (!(IN5)))) | IN8)) & ((!((((!(IN2)) & (!(IN1))) & IN3) & (!(IN5)))) | IN11)) & ((!(((IN2 & (!(IN1))) & IN3) & (!(IN5)))) | IN4)) & ((!((((!(IN2)) & IN1) & IN3) & (!(IN5)))) | IN13)) & ((!(((IN2 & IN1) & IN3) & (!(IN5)))) | IN10)) & ((!((((!(IN2)) & (!(IN1))) & (!(IN3))) & IN5)) | IN12)) & ((!(((IN2 & (!(IN1))) & (!(IN3))) & IN5)) | IN18)) & ((!((((!(IN2)) & IN1) & (!(IN3))) & IN5)) | IN16)) & ((!(((IN2 & IN1) & (!(IN3))) & IN5)) | IN14)) & ((!((((!(IN2)) & (!(IN1))) & IN3) & IN5)) | IN15)) & ((!(((IN2 & (!(IN1))) & IN3) & IN5)) | IN17)) & ((!((((!(IN2)) & IN1) & IN3) & IN5)) | IN19)) & ((!(((IN2 & IN1) & IN3) & IN5)) | IN20)

*)

FUNCTION_BLOCK F_CollectInput
  VAR_IN_OUT
      Data : ARRAY[1..20] OF BOOL;
  END_VAR
  VAR_INPUT
      TICK  : BOOL := 0;
      IN1   : BOOL := 0;
      IN2   : BOOL := 0;
      IN3   : BOOL := 0;
      IN4   : BOOL := 0;
      IN5   : BOOL := 0;
      RESET : BOOL := FALSE;
  END_VAR
  VAR_OUTPUT
      Finished : BOOL;
  END_VAR
  VAR
      j    : USINT := 1;
      tock : BOOL  := 0;
  END_VAR
  IF NOT RESET AND tock = NOT TICK THEN
      Data[j]   := IN1;
      Data[j+1] := IN2;
      Data[j+2] := IN3;
      Data[j+3] := IN4;
      Data[j+4] := IN5;
      j := j + 5;
      tock := TICK;
  ELSE
      j := 1;
      tock := 0;
  END_IF;
  Finished := (j > 20);
END_FUNCTION_BLOCK

PROGRAM Boiler
  VAR
    Data  : ARRAY[1..20] OF BOOL;
    Ready : BOOL;
    CollectInput : F_CollectInput;
  END_VAR
  VAR
    TICK     AT %IX1.0 : BOOL;
    IN1      AT %IX0.3 : BOOL;
    IN2      AT %IX0.4 : BOOL;
    IN3      AT %IX0.5 : BOOL;
    IN4      AT %IX0.6 : BOOL;
    IN5      AT %IX0.7 : BOOL;
    OutReady AT %QX0.0 : BOOL := FALSE;
    FeedNext AT %QX0.1 : BOOL := FALSE;
    Out      AT %QX0.2 : BOOL;
  END_VAR
  CollectInput(TICK:=TICK, IN1:=IN1, IN2:=IN2, IN3:=IN3, IN4:=IN4, IN5:=IN5);
  Ready := CollectInput.Finished;
  FeedNext := 1;
  IF Ready THEN
    Out := (((((((((((((((((NOT ((((NOT Data[2]) AND (NOT Data[1])) AND (NOT Data[3])) AND (NOT Data[5]))) OR Data[6]) AND ((NOT (((Data[2] AND (NOT Data[1])) AND (NOT Data[3])) AND (NOT Data[5]))) OR Data[7])) AND ((NOT ((((NOT Data[2]) AND Data[1]) AND (NOT Data[3])) AND (NOT Data[5]))) OR Data[9])) AND ((NOT (((Data[2] AND Data[1]) AND (NOT Data[3])) AND (NOT Data[5]))) OR Data[8])) AND ((NOT ((((NOT Data[2]) AND (NOT Data[1])) AND Data[3]) AND (NOT Data[5]))) OR Data[11])) AND ((NOT (((Data[2] AND (NOT Data[1])) AND Data[3]) AND (NOT Data[5]))) OR Data[4])) AND ((NOT ((((NOT Data[2]) AND Data[1]) AND Data[3]) AND (NOT Data[5]))) OR Data[13])) AND ((NOT (((Data[2] AND Data[1]) AND Data[3]) AND (NOT Data[5]))) OR Data[10])) AND ((NOT ((((NOT Data[2]) AND (NOT Data[1])) AND (NOT Data[3])) AND Data[5])) OR Data[12])) AND ((NOT (((Data[2] AND (NOT Data[1])) AND (NOT Data[3])) AND Data[5])) OR Data[18])) AND ((NOT ((((NOT Data[2]) AND Data[1]) AND (NOT Data[3])) AND Data[5])) OR Data[16])) AND ((NOT (((Data[2] AND Data[1]) AND (NOT Data[3])) AND Data[5])) OR Data[14])) AND ((NOT ((((NOT Data[2]) AND (NOT Data[1])) AND Data[3]) AND Data[5])) OR Data[15])) AND ((NOT (((Data[2] AND (NOT Data[1])) AND Data[3]) AND Data[5])) OR Data[17])) AND ((NOT ((((NOT Data[2]) AND Data[1]) AND Data[3]) AND Data[5])) OR Data[19])) AND ((NOT (((Data[2] AND Data[1]) AND Data[3]) AND Data[5])) OR Data[20]));
    OutReady := 1;
    CollectInput(RESET:=TRUE);
  END_IF;
END_PROGRAM

CONFIGURATION Config0
  RESOURCE Res0 ON PLC
    TASK task0(INTERVAL := T#20ms,PRIORITY := 0);
    PROGRAM instance0 WITH task0 : Boiler;
  END_RESOURCE
END_CONFIGURATION

(* ---- 4-MUX_whine-grads-sight.st ---- *)
(*
This code implements a shuffled multiplexer with 4 control bits.
The control bits are: Data[N3], Data[N1], Data[N2], Data[N4]
The input bits are: Data[N7], Data[N10], Data[N6], Data[N8], Data[N17], Data[N5], Data[N16], Data[N12], Data[N11], Data[N9], Data[N13], Data[N15], Data[N18], Data[N19], Data[N14], Data[N20]

The symbolic expression is:
((((((((((((((((!((((!(IN3)) & (!(IN1))) & (!(IN2))) & (!(IN4)))) | IN7) & ((!(((IN3 & (!(IN1))) & (!(IN2))) & (!(IN4)))) | IN10)) & ((!((((!(IN3)) & IN1) & (!(IN2))) & (!(IN4)))) | IN6)) & ((!(((IN3 & IN1) & (!(IN2))) & (!(IN4)))) | IN8)) & ((!((((!(IN3)) & (!(IN1))) & IN2) & (!(IN4)))) | IN17)) & ((!(((IN3 & (!(IN1))) & IN2) & (!(IN4)))) | IN5)) & ((!((((!(IN3)) & IN1) & IN2) & (!(IN4)))) | IN16)) & ((!(((IN3 & IN1) & IN2) & (!(IN4)))) | IN12)) & ((!((((!(IN3)) & (!(IN1))) & (!(IN2))) & IN4)) | IN11)) & ((!(((IN3 & (!(IN1))) & (!(IN2))) & IN4)) | IN9)) & ((!((((!(IN3)) & IN1) & (!(IN2))) & IN4)) | IN13)) & ((!(((IN3 & IN1) & (!(IN2))) & IN4)) | IN15)) & ((!((((!(IN3)) & (!(IN1))) & IN2) & IN4)) | IN18)) & ((!(((IN3 & (!(IN1))) & IN2) & IN4)) | IN19)) & ((!((((!(IN3)) & IN1) & IN2) & IN4)) | IN14)) & ((!(((IN3 & IN1) & IN2) & IN4)) | IN20)

*)

FUNCTION_BLOCK F_CollectInput
  VAR_IN_OUT
      Data : ARRAY[1..20] OF BOOL;
  END_VAR
  VAR_INPUT
      TICK  : BOOL := 0;
      IN1   : BOOL := 0;
      IN2   : BOOL := 0;
      IN3   : BOOL := 0;
      IN4   : BOOL := 0;
      IN5   : BOOL := 0;
      RESET : BOOL := FALSE;
  END_VAR
  VAR_OUTPUT
      Finished : BOOL;
  END_VAR
  VAR
      j    : USINT := 1;
      tock : BOOL  := 0;
  END_VAR
  IF NOT RESET AND tock = NOT TICK THEN
      Data[j]   := IN1;
      Data[j+1] := IN2;
      Data[j+2] := IN3;
      Data[j+3] := IN4;
      Data[j+4] := IN5;
      j := j + 5;
      tock := TICK;
  ELSE
      j := 1;
      tock := 0;
  END_IF;
  Finished := (j > 20);
END_FUNCTION_BLOCK

PROGRAM Boiler
  VAR
    Data  : ARRAY[1..20] OF BOOL;
    Ready : BOOL;
    CollectInput : F_CollectInput;
  END_VAR
  VAR
    TICK     AT %IX1.0 : BOOL;
    IN1      AT %IX0.3 : BOOL;
    IN2      AT %IX0.4 : BOOL;
    IN3      AT %IX0.5 : BOOL;
    IN4      AT %IX0.6 : BOOL;
    IN5      AT %IX0.7 : BOOL;
    OutReady AT %QX0.0 : BOOL := FALSE;
    FeedNext AT %QX0.1 : BOOL := FALSE;
    Out      AT %QX0.2 : BOOL;
  END_VAR
  CollectInput(TICK:=TICK, IN1:=IN1, IN2:=IN2, IN3:=IN3, IN4:=IN4, IN5:=IN5);
  Ready := CollectInput.Finished;
  FeedNext := 1;
  IF Ready THEN
    Out := (((((((((((((((((NOT ((((NOT Data[3]) AND (NOT Data[1])) AND (NOT Data[2])) AND (NOT Data[4]))) OR Data[7]) AND ((NOT (((Data[3] AND (NOT Data[1])) AND (NOT Data[2])) AND (NOT Data[4]))) OR Data[10])) AND ((NOT ((((NOT Data[3]) AND Data[1]) AND (NOT Data[2])) AND (NOT Data[4]))) OR Data[6])) AND ((NOT (((Data[3] AND Data[1]) AND (NOT Data[2])) AND (NOT Data[4]))) OR Data[8])) AND ((NOT ((((NOT Data[3]) AND (NOT Data[1])) AND Data[2]) AND (NOT Data[4]))) OR Data[17])) AND ((NOT (((Data[3] AND (NOT Data[1])) AND Data[2]) AND (NOT Data[4]))) OR Data[5])) AND ((NOT ((((NOT Data[3]) AND Data[1]) AND Data[2]) AND (NOT Data[4]))) OR Data[16])) AND ((NOT (((Data[3] AND Data[1]) AND Data[2]) AND (NOT Data[4]))) OR Data[12])) AND ((NOT ((((NOT Data[3]) AND (NOT Data[1])) AND (NOT Data[2])) AND Data[4])) OR Data[11])) AND ((NOT (((Data[3] AND (NOT Data[1])) AND (NOT Data[2])) AND Data[4])) OR Data[9])) AND ((NOT ((((NOT Data[3]) AND Data[1]) AND (NOT Data[2])) AND Data[4])) OR Data[13])) AND ((NOT (((Data[3] AND Data[1]) AND (NOT Data[2])) AND Data[4])) OR Data[15])) AND ((NOT ((((NOT Data[3]) AND (NOT Data[1])) AND Data[2]) AND Data[4])) OR Data[18])) AND ((NOT (((Data[3] AND (NOT Data[1])) AND Data[2]) AND Data[4])) OR Data[19])) AND ((NOT ((((NOT Data[3]) AND Data[1]) AND Data[2]) AND Data[4])) OR Data[14])) AND ((NOT (((Data[3] AND Data[1]) AND Data[2]) AND Data[4])) OR Data[20]));
    OutReady := 1;
    CollectInput(RESET:=TRUE);
  END_IF;
END_PROGRAM

CONFIGURATION Config0
  RESOURCE Res0 ON PLC
    TASK task0(INTERVAL := T#20ms,PRIORITY := 0);
    PROGRAM instance0 WITH task0 : Boiler;
  END_RESOURCE
END_CONFIGURATION

(* ---- 4-MUX_whorl-fetus-stuff.st ---- *)
(*
This code implements a shuffled multiplexer with 4 control bits.
The control bits are: Data[N1], Data[N2], Data[N9], Data[N3]
The input bits are: Data[N4], Data[N5], Data[N6], Data[N10], Data[N7], Data[N8], Data[N12], Data[N11], Data[N17], Data[N13], Data[N14], Data[N16], Data[N15], Data[N18], Data[N20], Data[N19]

The symbolic expression is:
((((((((((((((((!((((!(IN1)) & (!(IN2))) & (!(IN9))) & (!(IN3)))) | IN4) & ((!(((IN1 & (!(IN2))) & (!(IN9))) & (!(IN3)))) | IN5)) & ((!((((!(IN1)) & IN2) & (!(IN9))) & (!(IN3)))) | IN6)) & ((!(((IN1 & IN2) & (!(IN9))) & (!(IN3)))) | IN10)) & ((!((((!(IN1)) & (!(IN2))) & IN9) & (!(IN3)))) | IN7)) & ((!(((IN1 & (!(IN2))) & IN9) & (!(IN3)))) | IN8)) & ((!((((!(IN1)) & IN2) & IN9) & (!(IN3)))) | IN12)) & ((!(((IN1 & IN2) & IN9) & (!(IN3)))) | IN11)) & ((!((((!(IN1)) & (!(IN2))) & (!(IN9))) & IN3)) | IN17)) & ((!(((IN1 & (!(IN2))) & (!(IN9))) & IN3)) | IN13)) & ((!((((!(IN1)) & IN2) & (!(IN9))) & IN3)) | IN14)) & ((!(((IN1 & IN2) & (!(IN9))) & IN3)) | IN16)) & ((!((((!(IN1)) & (!(IN2))) & IN9) & IN3)) | IN15)) & ((!(((IN1 & (!(IN2))) & IN9) & IN3)) | IN18)) & ((!((((!(IN1)) & IN2) & IN9) & IN3)) | IN20)) & ((!(((IN1 & IN2) & IN9) & IN3)) | IN19)

*)

FUNCTION_BLOCK F_CollectInput
  VAR_IN_OUT
      Data : ARRAY[1..20] OF BOOL;
  END_VAR
  VAR_INPUT
      TICK  : BOOL := 0;
      IN1   : BOOL := 0;
      IN2   : BOOL := 0;
      IN3   : BOOL := 0;
      IN4   : BOOL := 0;
      IN5   : BOOL := 0;
      RESET : BOOL := FALSE;
  END_VAR
  VAR_OUTPUT
      Finished : BOOL;
  END_VAR
  VAR
      j    : USINT := 1;
      tock : BOOL  := 0;
  END_VAR
  IF NOT RESET AND tock = NOT TICK THEN
      Data[j]   := IN1;
      Data[j+1] := IN2;
      Data[j+2] := IN3;
      Data[j+3] := IN4;
      Data[j+4] := IN5;
      j := j + 5;
      tock := TICK;
  ELSE
      j := 1;
      tock := 0;
  END_IF;
  Finished := (j > 20);
END_FUNCTION_BLOCK

PROGRAM Boiler
  VAR
    Data  : ARRAY[1..20] OF BOOL;
    Ready : BOOL;
    CollectInput : F_CollectInput;
  END_VAR
  VAR
    TICK     AT %IX1.0 : BOOL;
    IN1      AT %IX0.3 : BOOL;
    IN2      AT %IX0.4 : BOOL;
    IN3      AT %IX0.5 : BOOL;
    IN4      AT %IX0.6 : BOOL;
    IN5      AT %IX0.7 : BOOL;
    OutReady AT %QX0.0 : BOOL := FALSE;
    FeedNext AT %QX0.1 : BOOL := FALSE;
    Out      AT %QX0.2 : BOOL;
  END_VAR
  CollectInput(TICK:=TICK, IN1:=IN1, IN2:=IN2, IN3:=IN3, IN4:=IN4, IN5:=IN5);
  Ready := CollectInput.Finished;
  FeedNext := 1;
  IF Ready THEN
    Out := (((((((((((((((((NOT ((((NOT Data[1]) AND (NOT Data[2])) AND (NOT Data[9])) AND (NOT Data[3]))) OR Data[4]) AND ((NOT (((Data[1] AND (NOT Data[2])) AND (NOT Data[9])) AND (NOT Data[3]))) OR Data[5])) AND ((NOT ((((NOT Data[1]) AND Data[2]) AND (NOT Data[9])) AND (NOT Data[3]))) OR Data[6])) AND ((NOT (((Data[1] AND Data[2]) AND (NOT Data[9])) AND (NOT Data[3]))) OR Data[10])) AND ((NOT ((((NOT Data[1]) AND (NOT Data[2])) AND Data[9]) AND (NOT Data[3]))) OR Data[7])) AND ((NOT (((Data[1] AND (NOT Data[2])) AND Data[9]) AND (NOT Data[3]))) OR Data[8])) AND ((NOT ((((NOT Data[1]) AND Data[2]) AND Data[9]) AND (NOT Data[3]))) OR Data[12])) AND ((NOT (((Data[1] AND Data[2]) AND Data[9]) AND (NOT Data[3]))) OR Data[11])) AND ((NOT ((((NOT Data[1]) AND (NOT Data[2])) AND (NOT Data[9])) AND Data[3])) OR Data[17])) AND ((NOT (((Data[1] AND (NOT Data[2])) AND (NOT Data[9])) AND Data[3])) OR Data[13])) AND ((NOT ((((NOT Data[1]) AND Data[2]) AND (NOT Data[9])) AND Data[3])) OR Data[14])) AND ((NOT (((Data[1] AND Data[2]) AND (NOT Data[9])) AND Data[3])) OR Data[16])) AND ((NOT ((((NOT Data[1]) AND (NOT Data[2])) AND Data[9]) AND Data[3])) OR Data[15])) AND ((NOT (((Data[1] AND (NOT Data[2])) AND Data[9]) AND Data[3])) OR Data[18])) AND ((NOT ((((NOT Data[1]) AND Data[2]) AND Data[9]) AND Data[3])) OR Data[20])) AND ((NOT (((Data[1] AND Data[2]) AND Data[9]) AND Data[3])) OR Data[19]));
    OutReady := 1;
    CollectInput(RESET:=TRUE);
  END_IF;
END_PROGRAM

CONFIGURATION Config0
  RESOURCE Res0 ON PLC
    TASK task0(INTERVAL := T#20ms,PRIORITY := 0);
    PROGRAM instance0 WITH task0 : Boiler;
  END_RESOURCE
END_CONFIGURATION

(* ---- 4-MUX_yokel-sniff-tenon.st ---- *)
(*
This code implements a shuffled multiplexer with 4 control bits.
The control bits are: Data[N1], Data[N3], Data[N2], Data[N4]
The input bits are: Data[N5], Data[N11], Data[N6], Data[N9], Data[N7], Data[N12], Data[N10], Data[N8], Data[N13], Data[N14], Data[N16], Data[N18], Data[N15], Data[N20], Data[N17], Data[N19]

The symbolic expression is:
((((((((((((((((!((((!(IN1)) & (!(IN3))) & (!(IN2))) & (!(IN4)))) | IN5) & ((!(((IN1 & (!(IN3))) & (!(IN2))) & (!(IN4)))) | IN11)) & ((!((((!(IN1)) & IN3) & (!(IN2))) & (!(IN4)))) | IN6)) & ((!(((IN1 & IN3) & (!(IN2))) & (!(IN4)))) | IN9)) & ((!((((!(IN1)) & (!(IN3))) & IN2) & (!(IN4)))) | IN7)) & ((!(((IN1 & (!(IN3))) & IN2) & (!(IN4)))) | IN12)) & ((!((((!(IN1)) & IN3) & IN2) & (!(IN4)))) | IN10)) & ((!(((IN1 & IN3) & IN2) & (!(IN4)))) | IN8)) & ((!((((!(IN1)) & (!(IN3))) & (!(IN2))) & IN4)) | IN13)) & ((!(((IN1 & (!(IN3))) & (!(IN2))) & IN4)) | IN14)) & ((!((((!(IN1)) & IN3) & (!(IN2))) & IN4)) | IN16)) & ((!(((IN1 & IN3) & (!(IN2))) & IN4)) | IN18)) & ((!((((!(IN1)) & (!(IN3))) & IN2) & IN4)) | IN15)) & ((!(((IN1 & (!(IN3))) & IN2) & IN4)) | IN20)) & ((!((((!(IN1)) & IN3) & IN2) & IN4)) | IN17)) & ((!(((IN1 & IN3) & IN2) & IN4)) | IN19)

*)

FUNCTION_BLOCK F_CollectInput
  VAR_IN_OUT
      Data : ARRAY[1..20] OF BOOL;
  END_VAR
  VAR_INPUT
      TICK  : BOOL := 0;
      IN1   : BOOL := 0;
      IN2   : BOOL := 0;
      IN3   : BOOL := 0;
      IN4   : BOOL := 0;
      IN5   : BOOL := 0;
      RESET : BOOL := FALSE;
  END_VAR
  VAR_OUTPUT
      Finished : BOOL;
  END_VAR
  VAR
      j    : USINT := 1;
      tock : BOOL  := 0;
  END_VAR
  IF NOT RESET AND tock = NOT TICK THEN
      Data[j]   := IN1;
      Data[j+1] := IN2;
      Data[j+2] := IN3;
      Data[j+3] := IN4;
      Data[j+4] := IN5;
      j := j + 5;
      tock := TICK;
  ELSE
      j := 1;
      tock := 0;
  END_IF;
  Finished := (j > 20);
END_FUNCTION_BLOCK

PROGRAM Boiler
  VAR
    Data  : ARRAY[1..20] OF BOOL;
    Ready : BOOL;
    CollectInput : F_CollectInput;
  END_VAR
  VAR
    TICK     AT %IX1.0 : BOOL;
    IN1      AT %IX0.3 : BOOL;
    IN2      AT %IX0.4 : BOOL;
    IN3      AT %IX0.5 : BOOL;
    IN4      AT %IX0.6 : BOOL;
    IN5      AT %IX0.7 : BOOL;
    OutReady AT %QX0.0 : BOOL := FALSE;
    FeedNext AT %QX0.1 : BOOL := FALSE;
    Out      AT %QX0.2 : BOOL;
  END_VAR
  CollectInput(TICK:=TICK, IN1:=IN1, IN2:=IN2, IN3:=IN3, IN4:=IN4, IN5:=IN5);
  Ready := CollectInput.Finished;
  FeedNext := 1;
  IF Ready THEN
    Out := (((((((((((((((((NOT ((((NOT Data[1]) AND (NOT Data[3])) AND (NOT Data[2])) AND (NOT Data[4]))) OR Data[5]) AND ((NOT (((Data[1] AND (NOT Data[3])) AND (NOT Data[2])) AND (NOT Data[4]))) OR Data[11])) AND ((NOT ((((NOT Data[1]) AND Data[3]) AND (NOT Data[2])) AND (NOT Data[4]))) OR Data[6])) AND ((NOT (((Data[1] AND Data[3]) AND (NOT Data[2])) AND (NOT Data[4]))) OR Data[9])) AND ((NOT ((((NOT Data[1]) AND (NOT Data[3])) AND Data[2]) AND (NOT Data[4]))) OR Data[7])) AND ((NOT (((Data[1] AND (NOT Data[3])) AND Data[2]) AND (NOT Data[4]))) OR Data[12])) AND ((NOT ((((NOT Data[1]) AND Data[3]) AND Data[2]) AND (NOT Data[4]))) OR Data[10])) AND ((NOT (((Data[1] AND Data[3]) AND Data[2]) AND (NOT Data[4]))) OR Data[8])) AND ((NOT ((((NOT Data[1]) AND (NOT Data[3])) AND (NOT Data[2])) AND Data[4])) OR Data[13])) AND ((NOT (((Data[1] AND (NOT Data[3])) AND (NOT Data[2])) AND Data[4])) OR Data[14])) AND ((NOT ((((NOT Data[1]) AND Data[3]) AND (NOT Data[2])) AND Data[4])) OR Data[16])) AND ((NOT (((Data[1] AND Data[3]) AND (NOT Data[2])) AND Data[4])) OR Data[18])) AND ((NOT ((((NOT Data[1]) AND (NOT Data[3])) AND Data[2]) AND Data[4])) OR Data[15])) AND ((NOT (((Data[1] AND (NOT Data[3])) AND Data[2]) AND Data[4])) OR Data[20])) AND ((NOT ((((NOT Data[1]) AND Data[3]) AND Data[2]) AND Data[4])) OR Data[17])) AND ((NOT (((Data[1] AND Data[3]) AND Data[2]) AND Data[4])) OR Data[19]));
    OutReady := 1;
    CollectInput(RESET:=TRUE);
  END_IF;
END_PROGRAM

CONFIGURATION Config0
  RESOURCE Res0 ON PLC
    TASK task0(INTERVAL := T#20ms,PRIORITY := 0);
    PROGRAM instance0 WITH task0 : Boiler;
  END_RESOURCE
END_CONFIGURATION

(* ---- 4-MUX_yowls-blood-clock.st ---- *)
(*
This code implements a shuffled multiplexer with 4 control bits.
The control bits are: Data[N1], Data[N3], Data[N2], Data[N4]
The input bits are: Data[N5], Data[N6], Data[N8], Data[N9], Data[N7], Data[N11], Data[N12], Data[N10], Data[N14], Data[N13], Data[N18], Data[N15], Data[N16], Data[N19], Data[N17], Data[N20]

The symbolic expression is:
((((((((((((((((!((((!(IN1)) & (!(IN3))) & (!(IN2))) & (!(IN4)))) | IN5) & ((!(((IN1 & (!(IN3))) & (!(IN2))) & (!(IN4)))) | IN6)) & ((!((((!(IN1)) & IN3) & (!(IN2))) & (!(IN4)))) | IN8)) & ((!(((IN1 & IN3) & (!(IN2))) & (!(IN4)))) | IN9)) & ((!((((!(IN1)) & (!(IN3))) & IN2) & (!(IN4)))) | IN7)) & ((!(((IN1 & (!(IN3))) & IN2) & (!(IN4)))) | IN11)) & ((!((((!(IN1)) & IN3) & IN2) & (!(IN4)))) | IN12)) & ((!(((IN1 & IN3) & IN2) & (!(IN4)))) | IN10)) & ((!((((!(IN1)) & (!(IN3))) & (!(IN2))) & IN4)) | IN14)) & ((!(((IN1 & (!(IN3))) & (!(IN2))) & IN4)) | IN13)) & ((!((((!(IN1)) & IN3) & (!(IN2))) & IN4)) | IN18)) & ((!(((IN1 & IN3) & (!(IN2))) & IN4)) | IN15)) & ((!((((!(IN1)) & (!(IN3))) & IN2) & IN4)) | IN16)) & ((!(((IN1 & (!(IN3))) & IN2) & IN4)) | IN19)) & ((!((((!(IN1)) & IN3) & IN2) & IN4)) | IN17)) & ((!(((IN1 & IN3) & IN2) & IN4)) | IN20)

*)

FUNCTION_BLOCK F_CollectInput
  VAR_IN_OUT
      Data : ARRAY[1..20] OF BOOL;
  END_VAR
  VAR_INPUT
      TICK  : BOOL := 0;
      IN1   : BOOL := 0;
      IN2   : BOOL := 0;
      IN3   : BOOL := 0;
      IN4   : BOOL := 0;
      IN5   : BOOL := 0;
      RESET : BOOL := FALSE;
  END_VAR
  VAR_OUTPUT
      Finished : BOOL;
  END_VAR
  VAR
      j    : USINT := 1;
      tock : BOOL  := 0;
  END_VAR
  IF NOT RESET AND tock = NOT TICK THEN
      Data[j]   := IN1;
      Data[j+1] := IN2;
      Data[j+2] := IN3;
      Data[j+3] := IN4;
      Data[j+4] := IN5;
      j := j + 5;
      tock := TICK;
  ELSE
      j := 1;
      tock := 0;
  END_IF;
  Finished := (j > 20);
END_FUNCTION_BLOCK

PROGRAM Boiler
  VAR
    Data  : ARRAY[1..20] OF BOOL;
    Ready : BOOL;
    CollectInput : F_CollectInput;
  END_VAR
  VAR
    TICK     AT %IX1.0 : BOOL;
    IN1      AT %IX0.3 : BOOL;
    IN2      AT %IX0.4 : BOOL;
    IN3      AT %IX0.5 : BOOL;
    IN4      AT %IX0.6 : BOOL;
    IN5      AT %IX0.7 : BOOL;
    OutReady AT %QX0.0 : BOOL := FALSE;
    FeedNext AT %QX0.1 : BOOL := FALSE;
    Out      AT %QX0.2 : BOOL;
  END_VAR
  CollectInput(TICK:=TICK, IN1:=IN1, IN2:=IN2, IN3:=IN3, IN4:=IN4, IN5:=IN5);
  Ready := CollectInput.Finished;
  FeedNext := 1;
  IF Ready THEN
    Out := (((((((((((((((((NOT ((((NOT Data[1]) AND (NOT Data[3])) AND (NOT Data[2])) AND (NOT Data[4]))) OR Data[5]) AND ((NOT (((Data[1] AND (NOT Data[3])) AND (NOT Data[2])) AND (NOT Data[4]))) OR Data[6])) AND ((NOT ((((NOT Data[1]) AND Data[3]) AND (NOT Data[2])) AND (NOT Data[4]))) OR Data[8])) AND ((NOT (((Data[1] AND Data[3]) AND (NOT Data[2])) AND (NOT Data[4]))) OR Data[9])) AND ((NOT ((((NOT Data[1]) AND (NOT Data[3])) AND Data[2]) AND (NOT Data[4]))) OR Data[7])) AND ((NOT (((Data[1] AND (NOT Data[3])) AND Data[2]) AND (NOT Data[4]))) OR Data[11])) AND ((NOT ((((NOT Data[1]) AND Data[3]) AND Data[2]) AND (NOT Data[4]))) OR Data[12])) AND ((NOT (((Data[1] AND Data[3]) AND Data[2]) AND (NOT Data[4]))) OR Data[10])) AND ((NOT ((((NOT Data[1]) AND (NOT Data[3])) AND (NOT Data[2])) AND Data[4])) OR Data[14])) AND ((NOT (((Data[1] AND (NOT Data[3])) AND (NOT Data[2])) AND Data[4])) OR Data[13])) AND ((NOT ((((NOT Data[1]) AND Data[3]) AND (NOT Data[2])) AND Data[4])) OR Data[18])) AND ((NOT (((Data[1] AND Data[3]) AND (NOT Data[2])) AND Data[4])) OR Data[15])) AND ((NOT ((((NOT Data[1]) AND (NOT Data[3])) AND Data[2]) AND Data[4])) OR Data[16])) AND ((NOT (((Data[1] AND (NOT Data[3])) AND Data[2]) AND Data[4])) OR Data[19])) AND ((NOT ((((NOT Data[1]) AND Data[3]) AND Data[2]) AND Data[4])) OR Data[17])) AND ((NOT (((Data[1] AND Data[3]) AND Data[2]) AND Data[4])) OR Data[20]));
    OutReady := 1;
    CollectInput(RESET:=TRUE);
  END_IF;
END_PROGRAM

CONFIGURATION Config0
  RESOURCE Res0 ON PLC
    TASK task0(INTERVAL := T#20ms,PRIORITY := 0);
    PROGRAM instance0 WITH task0 : Boiler;
  END_RESOURCE
END_CONFIGURATION

(* ---- 5-MUX_agley-purse-north.st ---- *)
(*
This code implements a shuffled multiplexer with 5 control bits.
The control bits are: Data[N3], Data[N5], Data[N21], Data[N23], Data[N20]
The input bits are: Data[N24], Data[N1], Data[N2], Data[N4], Data[N6], Data[N7], Data[N22], Data[N9], Data[N11], Data[N12], Data[N25], Data[N8], Data[N26], Data[N10], Data[N14], Data[N13], Data[N17], Data[N15], Data[N16], Data[N31], Data[N19], Data[N18], Data[N28], Data[N27], Data[N29], Data[N30], Data[N32], Data[N33], Data[N36], Data[N34], Data[N35], Data[N37]

The symbolic expression is:
((((((((((((((((((((((((((((((((!(((((!(IN3)) & (!(IN5))) & (!(IN21))) & (!(IN23))) & (!(IN20)))) | IN24) & ((!((((IN3 & (!(IN5))) & (!(IN21))) & (!(IN23))) & (!(IN20)))) | IN1)) & ((!(((((!(IN3)) & IN5) & (!(IN21))) & (!(IN23))) & (!(IN20)))) | IN2)) & ((!((((IN3 & IN5) & (!(IN21))) & (!(IN23))) & (!(IN20)))) | IN4)) & ((!(((((!(IN3)) & (!(IN5))) & IN21) & (!(IN23))) & (!(IN20)))) | IN6)) & ((!((((IN3 & (!(IN5))) & IN21) & (!(IN23))) & (!(IN20)))) | IN7)) & ((!(((((!(IN3)) & IN5) & IN21) & (!(IN23))) & (!(IN20)))) | IN22)) & ((!((((IN3 & IN5) & IN21) & (!(IN23))) & (!(IN20)))) | IN9)) & ((!(((((!(IN3)) & (!(IN5))) & (!(IN21))) & IN23) & (!(IN20)))) | IN11)) & ((!((((IN3 & (!(IN5))) & (!(IN21))) & IN23) & (!(IN20)))) | IN12)) & ((!(((((!(IN3)) & IN5) & (!(IN21))) & IN23) & (!(IN20)))) | IN25)) & ((!((((IN3 & IN5) & (!(IN21))) & IN23) & (!(IN20)))) | IN8)) & ((!(((((!(IN3)) & (!(IN5))) & IN21) & IN23) & (!(IN20)))) | IN26)) & ((!((((IN3 & (!(IN5))) & IN21) & IN23) & (!(IN20)))) | IN10)) & ((!(((((!(IN3)) & IN5) & IN21) & IN23) & (!(IN20)))) | IN14)) & ((!((((IN3 & IN5) & IN21) & IN23) & (!(IN20)))) | IN13)) & ((!(((((!(IN3)) & (!(IN5))) & (!(IN21))) & (!(IN23))) & IN20)) | IN17)) & ((!((((IN3 & (!(IN5))) & (!(IN21))) & (!(IN23))) & IN20)) | IN15)) & ((!(((((!(IN3)) & IN5) & (!(IN21))) & (!(IN23))) & IN20)) | IN16)) & ((!((((IN3 & IN5) & (!(IN21))) & (!(IN23))) & IN20)) | IN31)) & ((!(((((!(IN3)) & (!(IN5))) & IN21) & (!(IN23))) & IN20)) | IN19)) & ((!((((IN3 & (!(IN5))) & IN21) & (!(IN23))) & IN20)) | IN18)) & ((!(((((!(IN3)) & IN5) & IN21) & (!(IN23))) & IN20)) | IN28)) & ((!((((IN3 & IN5) & IN21) & (!(IN23))) & IN20)) | IN27)) & ((!(((((!(IN3)) & (!(IN5))) & (!(IN21))) & IN23) & IN20)) | IN29)) & ((!((((IN3 & (!(IN5))) & (!(IN21))) & IN23) & IN20)) | IN30)) & ((!(((((!(IN3)) & IN5) & (!(IN21))) & IN23) & IN20)) | IN32)) & ((!((((IN3 & IN5) & (!(IN21))) & IN23) & IN20)) | IN33)) & ((!(((((!(IN3)) & (!(IN5))) & IN21) & IN23) & IN20)) | IN36)) & ((!((((IN3 & (!(IN5))) & IN21) & IN23) & IN20)) | IN34)) & ((!(((((!(IN3)) & IN5) & IN21) & IN23) & IN20)) | IN35)) & ((!((((IN3 & IN5) & IN21) & IN23) & IN20)) | IN37)

*)

FUNCTION_BLOCK F_CollectInput
  VAR_IN_OUT
      Data : ARRAY[1..40] OF BOOL;
  END_VAR
  VAR_INPUT
      TICK  : BOOL := 0;
      IN1   : BOOL := 0;
      IN2   : BOOL := 0;
      IN3   : BOOL := 0;
      IN4   : BOOL := 0;
      IN5   : BOOL := 0;
      RESET : BOOL := FALSE;
  END_VAR
  VAR_OUTPUT
      Finished : BOOL;
  END_VAR
  VAR
      j    : USINT := 1;
      tock : BOOL  := 0;
  END_VAR
  IF NOT RESET AND tock = NOT TICK THEN
      Data[j]   := IN1;
      Data[j+1] := IN2;
      Data[j+2] := IN3;
      Data[j+3] := IN4;
      Data[j+4] := IN5;
      j := j + 5;
      tock := TICK;
  ELSE
      j := 1;
      tock := 0;
  END_IF;
  Finished := (j > 40);
END_FUNCTION_BLOCK

PROGRAM Boiler
  VAR
    Data  : ARRAY[1..40] OF BOOL;
    Ready : BOOL;
    CollectInput : F_CollectInput;
  END_VAR
  VAR
    TICK     AT %IX1.0 : BOOL;
    IN1      AT %IX0.3 : BOOL;
    IN2      AT %IX0.4 : BOOL;
    IN3      AT %IX0.5 : BOOL;
    IN4      AT %IX0.6 : BOOL;
    IN5      AT %IX0.7 : BOOL;
    OutReady AT %QX0.0 : BOOL := FALSE;
    FeedNext AT %QX0.1 : BOOL := FALSE;
    Out      AT %QX0.2 : BOOL;
  END_VAR
  CollectInput(TICK:=TICK, IN1:=IN1, IN2:=IN2, IN3:=IN3, IN4:=IN4, IN5:=IN5);
  Ready := CollectInput.Finished;
  FeedNext := 1;
  IF Ready THEN
    Out := (((((((((((((((((((((((((((((((((NOT (((((NOT Data[3]) AND (NOT Data[5])) AND (NOT Data[21])) AND (NOT Data[23])) AND (NOT Data[20]))) OR Data[24]) AND ((NOT ((((Data[3] AND (NOT Data[5])) AND (NOT Data[21])) AND (NOT Data[23])) AND (NOT Data[20]))) OR Data[1])) AND ((NOT (((((NOT Data[3]) AND Data[5]) AND (NOT Data[21])) AND (NOT Data[23])) AND (NOT Data[20]))) OR Data[2])) AND ((NOT ((((Data[3] AND Data[5]) AND (NOT Data[21])) AND (NOT Data[23])) AND (NOT Data[20]))) OR Data[4])) AND ((NOT (((((NOT Data[3]) AND (NOT Data[5])) AND Data[21]) AND (NOT Data[23])) AND (NOT Data[20]))) OR Data[6])) AND ((NOT ((((Data[3] AND (NOT Data[5])) AND Data[21]) AND (NOT Data[23])) AND (NOT Data[20]))) OR Data[7])) AND ((NOT (((((NOT Data[3]) AND Data[5]) AND Data[21]) AND (NOT Data[23])) AND (NOT Data[20]))) OR Data[22])) AND ((NOT ((((Data[3] AND Data[5]) AND Data[21]) AND (NOT Data[23])) AND (NOT Data[20]))) OR Data[9])) AND ((NOT (((((NOT Data[3]) AND (NOT Data[5])) AND (NOT Data[21])) AND Data[23]) AND (NOT Data[20]))) OR Data[11])) AND ((NOT ((((Data[3] AND (NOT Data[5])) AND (NOT Data[21])) AND Data[23]) AND (NOT Data[20]))) OR Data[12])) AND ((NOT (((((NOT Data[3]) AND Data[5]) AND (NOT Data[21])) AND Data[23]) AND (NOT Data[20]))) OR Data[25])) AND ((NOT ((((Data[3] AND Data[5]) AND (NOT Data[21])) AND Data[23]) AND (NOT Data[20]))) OR Data[8])) AND ((NOT (((((NOT Data[3]) AND (NOT Data[5])) AND Data[21]) AND Data[23]) AND (NOT Data[20]))) OR Data[26])) AND ((NOT ((((Data[3] AND (NOT Data[5])) AND Data[21]) AND Data[23]) AND (NOT Data[20]))) OR Data[10])) AND ((NOT (((((NOT Data[3]) AND Data[5]) AND Data[21]) AND Data[23]) AND (NOT Data[20]))) OR Data[14])) AND ((NOT ((((Data[3] AND Data[5]) AND Data[21]) AND Data[23]) AND (NOT Data[20]))) OR Data[13])) AND ((NOT (((((NOT Data[3]) AND (NOT Data[5])) AND (NOT Data[21])) AND (NOT Data[23])) AND Data[20])) OR Data[17])) AND ((NOT ((((Data[3] AND (NOT Data[5])) AND (NOT Data[21])) AND (NOT Data[23])) AND Data[20])) OR Data[15])) AND ((NOT (((((NOT Data[3]) AND Data[5]) AND (NOT Data[21])) AND (NOT Data[23])) AND Data[20])) OR Data[16])) AND ((NOT ((((Data[3] AND Data[5]) AND (NOT Data[21])) AND (NOT Data[23])) AND Data[20])) OR Data[31])) AND ((NOT (((((NOT Data[3]) AND (NOT Data[5])) AND Data[21]) AND (NOT Data[23])) AND Data[20])) OR Data[19])) AND ((NOT ((((Data[3] AND (NOT Data[5])) AND Data[21]) AND (NOT Data[23])) AND Data[20])) OR Data[18])) AND ((NOT (((((NOT Data[3]) AND Data[5]) AND Data[21]) AND (NOT Data[23])) AND Data[20])) OR Data[28])) AND ((NOT ((((Data[3] AND Data[5]) AND Data[21]) AND (NOT Data[23])) AND Data[20])) OR Data[27])) AND ((NOT (((((NOT Data[3]) AND (NOT Data[5])) AND (NOT Data[21])) AND Data[23]) AND Data[20])) OR Data[29])) AND ((NOT ((((Data[3] AND (NOT Data[5])) AND (NOT Data[21])) AND Data[23]) AND Data[20])) OR Data[30])) AND ((NOT (((((NOT Data[3]) AND Data[5]) AND (NOT Data[21])) AND Data[23]) AND Data[20])) OR Data[32])) AND ((NOT ((((Data[3] AND Data[5]) AND (NOT Data[21])) AND Data[23]) AND Data[20])) OR Data[33])) AND ((NOT (((((NOT Data[3]) AND (NOT Data[5])) AND Data[21]) AND Data[23]) AND Data[20])) OR Data[36])) AND ((NOT ((((Data[3] AND (NOT Data[5])) AND Data[21]) AND Data[23]) AND Data[20])) OR Data[34])) AND ((NOT (((((NOT Data[3]) AND Data[5]) AND Data[21]) AND Data[23]) AND Data[20])) OR Data[35])) AND ((NOT ((((Data[3] AND Data[5]) AND Data[21]) AND Data[23]) AND Data[20])) OR Data[37]));
    OutReady := 1;
    CollectInput(RESET:=TRUE);
  END_IF;
END_PROGRAM

CONFIGURATION Config0
  RESOURCE Res0 ON PLC
    TASK task0(INTERVAL := T#20ms,PRIORITY := 0);
    PROGRAM instance0 WITH task0 : Boiler;
  END_RESOURCE
END_CONFIGURATION

(* ---- 5-MUX_alias-dieth-grant.st ---- *)
(*
This code implements a shuffled multiplexer with 5 control bits.
The control bits are: Data[N22], Data[N1], Data[N2], Data[N7], Data[N3]
The input bits are: Data[N5], Data[N4], Data[N20], Data[N11], Data[N21], Data[N8], Data[N23], Data[N9], Data[N26], Data[N12], Data[N24], Data[N27], Data[N6], Data[N25], Data[N28], Data[N10], Data[N13], Data[N16], Data[N17], Data[N29], Data[N14], Data[N15], Data[N30], Data[N32], Data[N31], Data[N35], Data[N18], Data[N19], Data[N33], Data[N34], Data[N36], Data[N37]

The symbolic expression is:
((((((((((((((((((((((((((((((((!(((((!(IN22)) & (!(IN1))) & (!(IN2))) & (!(IN7))) & (!(IN3)))) | IN5) & ((!((((IN22 & (!(IN1))) & (!(IN2))) & (!(IN7))) & (!(IN3)))) | IN4)) & ((!(((((!(IN22)) & IN1) & (!(IN2))) & (!(IN7))) & (!(IN3)))) | IN20)) & ((!((((IN22 & IN1) & (!(IN2))) & (!(IN7))) & (!(IN3)))) | IN11)) & ((!(((((!(IN22)) & (!(IN1))) & IN2) & (!(IN7))) & (!(IN3)))) | IN21)) & ((!((((IN22 & (!(IN1))) & IN2) & (!(IN7))) & (!(IN3)))) | IN8)) & ((!(((((!(IN22)) & IN1) & IN2) & (!(IN7))) & (!(IN3)))) | IN23)) & ((!((((IN22 & IN1) & IN2) & (!(IN7))) & (!(IN3)))) | IN9)) & ((!(((((!(IN22)) & (!(IN1))) & (!(IN2))) & IN7) & (!(IN3)))) | IN26)) & ((!((((IN22 & (!(IN1))) & (!(IN2))) & IN7) & (!(IN3)))) | IN12)) & ((!(((((!(IN22)) & IN1) & (!(IN2))) & IN7) & (!(IN3)))) | IN24)) & ((!((((IN22 & IN1) & (!(IN2))) & IN7) & (!(IN3)))) | IN27)) & ((!(((((!(IN22)) & (!(IN1))) & IN2) & IN7) & (!(IN3)))) | IN6)) & ((!((((IN22 & (!(IN1))) & IN2) & IN7) & (!(IN3)))) | IN25)) & ((!(((((!(IN22)) & IN1) & IN2) & IN7) & (!(IN3)))) | IN28)) & ((!((((IN22 & IN1) & IN2) & IN7) & (!(IN3)))) | IN10)) & ((!(((((!(IN22)) & (!(IN1))) & (!(IN2))) & (!(IN7))) & IN3)) | IN13)) & ((!((((IN22 & (!(IN1))) & (!(IN2))) & (!(IN7))) & IN3)) | IN16)) & ((!(((((!(IN22)) & IN1) & (!(IN2))) & (!(IN7))) & IN3)) | IN17)) & ((!((((IN22 & IN1) & (!(IN2))) & (!(IN7))) & IN3)) | IN29)) & ((!(((((!(IN22)) & (!(IN1))) & IN2) & (!(IN7))) & IN3)) | IN14)) & ((!((((IN22 & (!(IN1))) & IN2) & (!(IN7))) & IN3)) | IN15)) & ((!(((((!(IN22)) & IN1) & IN2) & (!(IN7))) & IN3)) | IN30)) & ((!((((IN22 & IN1) & IN2) & (!(IN7))) & IN3)) | IN32)) & ((!(((((!(IN22)) & (!(IN1))) & (!(IN2))) & IN7) & IN3)) | IN31)) & ((!((((IN22 & (!(IN1))) & (!(IN2))) & IN7) & IN3)) | IN35)) & ((!(((((!(IN22)) & IN1) & (!(IN2))) & IN7) & IN3)) | IN18)) & ((!((((IN22 & IN1) & (!(IN2))) & IN7) & IN3)) | IN19)) & ((!(((((!(IN22)) & (!(IN1))) & IN2) & IN7) & IN3)) | IN33)) & ((!((((IN22 & (!(IN1))) & IN2) & IN7) & IN3)) | IN34)) & ((!(((((!(IN22)) & IN1) & IN2) & IN7) & IN3)) | IN36)) & ((!((((IN22 & IN1) & IN2) & IN7) & IN3)) | IN37)

*)

FUNCTION_BLOCK F_CollectInput
  VAR_IN_OUT
      Data : ARRAY[1..40] OF BOOL;
  END_VAR
  VAR_INPUT
      TICK  : BOOL := 0;
      IN1   : BOOL := 0;
      IN2   : BOOL := 0;
      IN3   : BOOL := 0;
      IN4   : BOOL := 0;
      IN5   : BOOL := 0;
      RESET : BOOL := FALSE;
  END_VAR
  VAR_OUTPUT
      Finished : BOOL;
  END_VAR
  VAR
      j    : USINT := 1;
      tock : BOOL  := 0;
  END_VAR
  IF NOT RESET AND tock = NOT TICK THEN
      Data[j]   := IN1;
      Data[j+1] := IN2;
      Data[j+2] := IN3;
      Data[j+3] := IN4;
      Data[j+4] := IN5;
      j := j + 5;
      tock := TICK;
  ELSE
      j := 1;
      tock := 0;
  END_IF;
  Finished := (j > 40);
END_FUNCTION_BLOCK

PROGRAM Boiler
  VAR
    Data  : ARRAY[1..40] OF BOOL;
    Ready : BOOL;
    CollectInput : F_CollectInput;
  END_VAR
  VAR
    TICK     AT %IX1.0 : BOOL;
    IN1      AT %IX0.3 : BOOL;
    IN2      AT %IX0.4 : BOOL;
    IN3      AT %IX0.5 : BOOL;
    IN4      AT %IX0.6 : BOOL;
    IN5      AT %IX0.7 : BOOL;
    OutReady AT %QX0.0 : BOOL := FALSE;
    FeedNext AT %QX0.1 : BOOL := FALSE;
    Out      AT %QX0.2 : BOOL;
  END_VAR
  CollectInput(TICK:=TICK, IN1:=IN1, IN2:=IN2, IN3:=IN3, IN4:=IN4, IN5:=IN5);
  Ready := CollectInput.Finished;
  FeedNext := 1;
  IF Ready THEN
    Out := (((((((((((((((((((((((((((((((((NOT (((((NOT Data[22]) AND (NOT Data[1])) AND (NOT Data[2])) AND (NOT Data[7])) AND (NOT Data[3]))) OR Data[5]) AND ((NOT ((((Data[22] AND (NOT Data[1])) AND (NOT Data[2])) AND (NOT Data[7])) AND (NOT Data[3]))) OR Data[4])) AND ((NOT (((((NOT Data[22]) AND Data[1]) AND (NOT Data[2])) AND (NOT Data[7])) AND (NOT Data[3]))) OR Data[20])) AND ((NOT ((((Data[22] AND Data[1]) AND (NOT Data[2])) AND (NOT Data[7])) AND (NOT Data[3]))) OR Data[11])) AND ((NOT (((((NOT Data[22]) AND (NOT Data[1])) AND Data[2]) AND (NOT Data[7])) AND (NOT Data[3]))) OR Data[21])) AND ((NOT ((((Data[22] AND (NOT Data[1])) AND Data[2]) AND (NOT Data[7])) AND (NOT Data[3]))) OR Data[8])) AND ((NOT (((((NOT Data[22]) AND Data[1]) AND Data[2]) AND (NOT Data[7])) AND (NOT Data[3]))) OR Data[23])) AND ((NOT ((((Data[22] AND Data[1]) AND Data[2]) AND (NOT Data[7])) AND (NOT Data[3]))) OR Data[9])) AND ((NOT (((((NOT Data[22]) AND (NOT Data[1])) AND (NOT Data[2])) AND Data[7]) AND (NOT Data[3]))) OR Data[26])) AND ((NOT ((((Data[22] AND (NOT Data[1])) AND (NOT Data[2])) AND Data[7]) AND (NOT Data[3]))) OR Data[12])) AND ((NOT (((((NOT Data[22]) AND Data[1]) AND (NOT Data[2])) AND Data[7]) AND (NOT Data[3]))) OR Data[24])) AND ((NOT ((((Data[22] AND Data[1]) AND (NOT Data[2])) AND Data[7]) AND (NOT Data[3]))) OR Data[27])) AND ((NOT (((((NOT Data[22]) AND (NOT Data[1])) AND Data[2]) AND Data[7]) AND (NOT Data[3]))) OR Data[6])) AND ((NOT ((((Data[22] AND (NOT Data[1])) AND Data[2]) AND Data[7]) AND (NOT Data[3]))) OR Data[25])) AND ((NOT (((((NOT Data[22]) AND Data[1]) AND Data[2]) AND Data[7]) AND (NOT Data[3]))) OR Data[28])) AND ((NOT ((((Data[22] AND Data[1]) AND Data[2]) AND Data[7]) AND (NOT Data[3]))) OR Data[10])) AND ((NOT (((((NOT Data[22]) AND (NOT Data[1])) AND (NOT Data[2])) AND (NOT Data[7])) AND Data[3])) OR Data[13])) AND ((NOT ((((Data[22] AND (NOT Data[1])) AND (NOT Data[2])) AND (NOT Data[7])) AND Data[3])) OR Data[16])) AND ((NOT (((((NOT Data[22]) AND Data[1]) AND (NOT Data[2])) AND (NOT Data[7])) AND Data[3])) OR Data[17])) AND ((NOT ((((Data[22] AND Data[1]) AND (NOT Data[2])) AND (NOT Data[7])) AND Data[3])) OR Data[29])) AND ((NOT (((((NOT Data[22]) AND (NOT Data[1])) AND Data[2]) AND (NOT Data[7])) AND Data[3])) OR Data[14])) AND ((NOT ((((Data[22] AND (NOT Data[1])) AND Data[2]) AND (NOT Data[7])) AND Data[3])) OR Data[15])) AND ((NOT (((((NOT Data[22]) AND Data[1]) AND Data[2]) AND (NOT Data[7])) AND Data[3])) OR Data[30])) AND ((NOT ((((Data[22] AND Data[1]) AND Data[2]) AND (NOT Data[7])) AND Data[3])) OR Data[32])) AND ((NOT (((((NOT Data[22]) AND (NOT Data[1])) AND (NOT Data[2])) AND Data[7]) AND Data[3])) OR Data[31])) AND ((NOT ((((Data[22] AND (NOT Data[1])) AND (NOT Data[2])) AND Data[7]) AND Data[3])) OR Data[35])) AND ((NOT (((((NOT Data[22]) AND Data[1]) AND (NOT Data[2])) AND Data[7]) AND Data[3])) OR Data[18])) AND ((NOT ((((Data[22] AND Data[1]) AND (NOT Data[2])) AND Data[7]) AND Data[3])) OR Data[19])) AND ((NOT (((((NOT Data[22]) AND (NOT Data[1])) AND Data[2]) AND Data[7]) AND Data[3])) OR Data[33])) AND ((NOT ((((Data[22] AND (NOT Data[1])) AND Data[2]) AND Data[7]) AND Data[3])) OR Data[34])) AND ((NOT (((((NOT Data[22]) AND Data[1]) AND Data[2]) AND Data[7]) AND Data[3])) OR Data[36])) AND ((NOT ((((Data[22] AND Data[1]) AND Data[2]) AND Data[7]) AND Data[3])) OR Data[37]));
    OutReady := 1;
    CollectInput(RESET:=TRUE);
  END_IF;
END_PROGRAM

CONFIGURATION Config0
  RESOURCE Res0 ON PLC
    TASK task0(INTERVAL := T#20ms,PRIORITY := 0);
    PROGRAM instance0 WITH task0 : Boiler;
  END_RESOURCE
END_CONFIGURATION

(* ---- 5-MUX_amahs-began-skoal.st ---- *)
(*
This code implements a shuffled multiplexer with 5 control bits.
The control bits are: Data[N20], Data[N4], Data[N1], Data[N2], Data[N22]
The input bits are: Data[N24], Data[N21], Data[N3], Data[N25], Data[N27], Data[N9], Data[N6], Data[N5], Data[N7], Data[N8], Data[N10], Data[N30], Data[N11], Data[N23], Data[N26], Data[N28], Data[N29], Data[N31], Data[N12], Data[N13], Data[N33], Data[N14], Data[N32], Data[N15], Data[N16], Data[N34], Data[N17], Data[N35], Data[N37], Data[N18], Data[N36], Data[N19]

The symbolic expression is:
((((((((((((((((((((((((((((((((!(((((!(IN20)) & (!(IN4))) & (!(IN1))) & (!(IN2))) & (!(IN22)))) | IN24) & ((!((((IN20 & (!(IN4))) & (!(IN1))) & (!(IN2))) & (!(IN22)))) | IN21)) & ((!(((((!(IN20)) & IN4) & (!(IN1))) & (!(IN2))) & (!(IN22)))) | IN3)) & ((!((((IN20 & IN4) & (!(IN1))) & (!(IN2))) & (!(IN22)))) | IN25)) & ((!(((((!(IN20)) & (!(IN4))) & IN1) & (!(IN2))) & (!(IN22)))) | IN27)) & ((!((((IN20 & (!(IN4))) & IN1) & (!(IN2))) & (!(IN22)))) | IN9)) & ((!(((((!(IN20)) & IN4) & IN1) & (!(IN2))) & (!(IN22)))) | IN6)) & ((!((((IN20 & IN4) & IN1) & (!(IN2))) & (!(IN22)))) | IN5)) & ((!(((((!(IN20)) & (!(IN4))) & (!(IN1))) & IN2) & (!(IN22)))) | IN7)) & ((!((((IN20 & (!(IN4))) & (!(IN1))) & IN2) & (!(IN22)))) | IN8)) & ((!(((((!(IN20)) & IN4) & (!(IN1))) & IN2) & (!(IN22)))) | IN10)) & ((!((((IN20 & IN4) & (!(IN1))) & IN2) & (!(IN22)))) | IN30)) & ((!(((((!(IN20)) & (!(IN4))) & IN1) & IN2) & (!(IN22)))) | IN11)) & ((!((((IN20 & (!(IN4))) & IN1) & IN2) & (!(IN22)))) | IN23)) & ((!(((((!(IN20)) & IN4) & IN1) & IN2) & (!(IN22)))) | IN26)) & ((!((((IN20 & IN4) & IN1) & IN2) & (!(IN22)))) | IN28)) & ((!(((((!(IN20)) & (!(IN4))) & (!(IN1))) & (!(IN2))) & IN22)) | IN29)) & ((!((((IN20 & (!(IN4))) & (!(IN1))) & (!(IN2))) & IN22)) | IN31)) & ((!(((((!(IN20)) & IN4) & (!(IN1))) & (!(IN2))) & IN22)) | IN12)) & ((!((((IN20 & IN4) & (!(IN1))) & (!(IN2))) & IN22)) | IN13)) & ((!(((((!(IN20)) & (!(IN4))) & IN1) & (!(IN2))) & IN22)) | IN33)) & ((!((((IN20 & (!(IN4))) & IN1) & (!(IN2))) & IN22)) | IN14)) & ((!(((((!(IN20)) & IN4) & IN1) & (!(IN2))) & IN22)) | IN32)) & ((!((((IN20 & IN4) & IN1) & (!(IN2))) & IN22)) | IN15)) & ((!(((((!(IN20)) & (!(IN4))) & (!(IN1))) & IN2) & IN22)) | IN16)) & ((!((((IN20 & (!(IN4))) & (!(IN1))) & IN2) & IN22)) | IN34)) & ((!(((((!(IN20)) & IN4) & (!(IN1))) & IN2) & IN22)) | IN17)) & ((!((((IN20 & IN4) & (!(IN1))) & IN2) & IN22)) | IN35)) & ((!(((((!(IN20)) & (!(IN4))) & IN1) & IN2) & IN22)) | IN37)) & ((!((((IN20 & (!(IN4))) & IN1) & IN2) & IN22)) | IN18)) & ((!(((((!(IN20)) & IN4) & IN1) & IN2) & IN22)) | IN36)) & ((!((((IN20 & IN4) & IN1) & IN2) & IN22)) | IN19)

*)

FUNCTION_BLOCK F_CollectInput
  VAR_IN_OUT
      Data : ARRAY[1..40] OF BOOL;
  END_VAR
  VAR_INPUT
      TICK  : BOOL := 0;
      IN1   : BOOL := 0;
      IN2   : BOOL := 0;
      IN3   : BOOL := 0;
      IN4   : BOOL := 0;
      IN5   : BOOL := 0;
      RESET : BOOL := FALSE;
  END_VAR
  VAR_OUTPUT
      Finished : BOOL;
  END_VAR
  VAR
      j    : USINT := 1;
      tock : BOOL  := 0;
  END_VAR
  IF NOT RESET AND tock = NOT TICK THEN
      Data[j]   := IN1;
      Data[j+1] := IN2;
      Data[j+2] := IN3;
      Data[j+3] := IN4;
      Data[j+4] := IN5;
      j := j + 5;
      tock := TICK;
  ELSE
      j := 1;
      tock := 0;
  END_IF;
  Finished := (j > 40);
END_FUNCTION_BLOCK

PROGRAM Boiler
  VAR
    Data  : ARRAY[1..40] OF BOOL;
    Ready : BOOL;
    CollectInput : F_CollectInput;
  END_VAR
  VAR
    TICK     AT %IX1.0 : BOOL;
    IN1      AT %IX0.3 : BOOL;
    IN2      AT %IX0.4 : BOOL;
    IN3      AT %IX0.5 : BOOL;
    IN4      AT %IX0.6 : BOOL;
    IN5      AT %IX0.7 : BOOL;
    OutReady AT %QX0.0 : BOOL := FALSE;
    FeedNext AT %QX0.1 : BOOL := FALSE;
    Out      AT %QX0.2 : BOOL;
  END_VAR
  CollectInput(TICK:=TICK, IN1:=IN1, IN2:=IN2, IN3:=IN3, IN4:=IN4, IN5:=IN5);
  Ready := CollectInput.Finished;
  FeedNext := 1;
  IF Ready THEN
    Out := (((((((((((((((((((((((((((((((((NOT (((((NOT Data[20]) AND (NOT Data[4])) AND (NOT Data[1])) AND (NOT Data[2])) AND (NOT Data[22]))) OR Data[24]) AND ((NOT ((((Data[20] AND (NOT Data[4])) AND (NOT Data[1])) AND (NOT Data[2])) AND (NOT Data[22]))) OR Data[21])) AND ((NOT (((((NOT Data[20]) AND Data[4]) AND (NOT Data[1])) AND (NOT Data[2])) AND (NOT Data[22]))) OR Data[3])) AND ((NOT ((((Data[20] AND Data[4]) AND (NOT Data[1])) AND (NOT Data[2])) AND (NOT Data[22]))) OR Data[25])) AND ((NOT (((((NOT Data[20]) AND (NOT Data[4])) AND Data[1]) AND (NOT Data[2])) AND (NOT Data[22]))) OR Data[27])) AND ((NOT ((((Data[20] AND (NOT Data[4])) AND Data[1]) AND (NOT Data[2])) AND (NOT Data[22]))) OR Data[9])) AND ((NOT (((((NOT Data[20]) AND Data[4]) AND Data[1]) AND (NOT Data[2])) AND (NOT Data[22]))) OR Data[6])) AND ((NOT ((((Data[20] AND Data[4]) AND Data[1]) AND (NOT Data[2])) AND (NOT Data[22]))) OR Data[5])) AND ((NOT (((((NOT Data[20]) AND (NOT Data[4])) AND (NOT Data[1])) AND Data[2]) AND (NOT Data[22]))) OR Data[7])) AND ((NOT ((((Data[20] AND (NOT Data[4])) AND (NOT Data[1])) AND Data[2]) AND (NOT Data[22]))) OR Data[8])) AND ((NOT (((((NOT Data[20]) AND Data[4]) AND (NOT Data[1])) AND Data[2]) AND (NOT Data[22]))) OR Data[10])) AND ((NOT ((((Data[20] AND Data[4]) AND (NOT Data[1])) AND Data[2]) AND (NOT Data[22]))) OR Data[30])) AND ((NOT (((((NOT Data[20]) AND (NOT Data[4])) AND Data[1]) AND Data[2]) AND (NOT Data[22]))) OR Data[11])) AND ((NOT ((((Data[20] AND (NOT Data[4])) AND Data[1]) AND Data[2]) AND (NOT Data[22]))) OR Data[23])) AND ((NOT (((((NOT Data[20]) AND Data[4]) AND Data[1]) AND Data[2]) AND (NOT Data[22]))) OR Data[26])) AND ((NOT ((((Data[20] AND Data[4]) AND Data[1]) AND Data[2]) AND (NOT Data[22]))) OR Data[28])) AND ((NOT (((((NOT Data[20]) AND (NOT Data[4])) AND (NOT Data[1])) AND (NOT Data[2])) AND Data[22])) OR Data[29])) AND ((NOT ((((Data[20] AND (NOT Data[4])) AND (NOT Data[1])) AND (NOT Data[2])) AND Data[22])) OR Data[31])) AND ((NOT (((((NOT Data[20]) AND Data[4]) AND (NOT Data[1])) AND (NOT Data[2])) AND Data[22])) OR Data[12])) AND ((NOT ((((Data[20] AND Data[4]) AND (NOT Data[1])) AND (NOT Data[2])) AND Data[22])) OR Data[13])) AND ((NOT (((((NOT Data[20]) AND (NOT Data[4])) AND Data[1]) AND (NOT Data[2])) AND Data[22])) OR Data[33])) AND ((NOT ((((Data[20] AND (NOT Data[4])) AND Data[1]) AND (NOT Data[2])) AND Data[22])) OR Data[14])) AND ((NOT (((((NOT Data[20]) AND Data[4]) AND Data[1]) AND (NOT Data[2])) AND Data[22])) OR Data[32])) AND ((NOT ((((Data[20] AND Data[4]) AND Data[1]) AND (NOT Data[2])) AND Data[22])) OR Data[15])) AND ((NOT (((((NOT Data[20]) AND (NOT Data[4])) AND (NOT Data[1])) AND Data[2]) AND Data[22])) OR Data[16])) AND ((NOT ((((Data[20] AND (NOT Data[4])) AND (NOT Data[1])) AND Data[2]) AND Data[22])) OR Data[34])) AND ((NOT (((((NOT Data[20]) AND Data[4]) AND (NOT Data[1])) AND Data[2]) AND Data[22])) OR Data[17])) AND ((NOT ((((Data[20] AND Data[4]) AND (NOT Data[1])) AND Data[2]) AND Data[22])) OR Data[35])) AND ((NOT (((((NOT Data[20]) AND (NOT Data[4])) AND Data[1]) AND Data[2]) AND Data[22])) OR Data[37])) AND ((NOT ((((Data[20] AND (NOT Data[4])) AND Data[1]) AND Data[2]) AND Data[22])) OR Data[18])) AND ((NOT (((((NOT Data[20]) AND Data[4]) AND Data[1]) AND Data[2]) AND Data[22])) OR Data[36])) AND ((NOT ((((Data[20] AND Data[4]) AND Data[1]) AND Data[2]) AND Data[22])) OR Data[19]));
    OutReady := 1;
    CollectInput(RESET:=TRUE);
  END_IF;
END_PROGRAM

CONFIGURATION Config0
  RESOURCE Res0 ON PLC
    TASK task0(INTERVAL := T#20ms,PRIORITY := 0);
    PROGRAM instance0 WITH task0 : Boiler;
  END_RESOURCE
END_CONFIGURATION

(* ---- 5-MUX_amine-rived-hurts.st ---- *)
(*
This code implements a shuffled multiplexer with 5 control bits.
The control bits are: Data[N1], Data[N22], Data[N2], Data[N3], Data[N21]
The input bits are: Data[N23], Data[N5], Data[N4], Data[N6], Data[N8], Data[N20], Data[N24], Data[N26], Data[N25], Data[N27], Data[N13], Data[N11], Data[N9], Data[N15], Data[N31], Data[N28], Data[N29], Data[N33], Data[N14], Data[N7], Data[N32], Data[N18], Data[N30], Data[N10], Data[N17], Data[N36], Data[N16], Data[N19], Data[N12], Data[N34], Data[N37], Data[N35]

The symbolic expression is:
((((((((((((((((((((((((((((((((!(((((!(IN1)) & (!(IN22))) & (!(IN2))) & (!(IN3))) & (!(IN21)))) | IN23) & ((!((((IN1 & (!(IN22))) & (!(IN2))) & (!(IN3))) & (!(IN21)))) | IN5)) & ((!(((((!(IN1)) & IN22) & (!(IN2))) & (!(IN3))) & (!(IN21)))) | IN4)) & ((!((((IN1 & IN22) & (!(IN2))) & (!(IN3))) & (!(IN21)))) | IN6)) & ((!(((((!(IN1)) & (!(IN22))) & IN2) & (!(IN3))) & (!(IN21)))) | IN8)) & ((!((((IN1 & (!(IN22))) & IN2) & (!(IN3))) & (!(IN21)))) | IN20)) & ((!(((((!(IN1)) & IN22) & IN2) & (!(IN3))) & (!(IN21)))) | IN24)) & ((!((((IN1 & IN22) & IN2) & (!(IN3))) & (!(IN21)))) | IN26)) & ((!(((((!(IN1)) & (!(IN22))) & (!(IN2))) & IN3) & (!(IN21)))) | IN25)) & ((!((((IN1 & (!(IN22))) & (!(IN2))) & IN3) & (!(IN21)))) | IN27)) & ((!(((((!(IN1)) & IN22) & (!(IN2))) & IN3) & (!(IN21)))) | IN13)) & ((!((((IN1 & IN22) & (!(IN2))) & IN3) & (!(IN21)))) | IN11)) & ((!(((((!(IN1)) & (!(IN22))) & IN2) & IN3) & (!(IN21)))) | IN9)) & ((!((((IN1 & (!(IN22))) & IN2) & IN3) & (!(IN21)))) | IN15)) & ((!(((((!(IN1)) & IN22) & IN2) & IN3) & (!(IN21)))) | IN31)) & ((!((((IN1 & IN22) & IN2) & IN3) & (!(IN21)))) | IN28)) & ((!(((((!(IN1)) & (!(IN22))) & (!(IN2))) & (!(IN3))) & IN21)) | IN29)) & ((!((((IN1 & (!(IN22))) & (!(IN2))) & (!(IN3))) & IN21)) | IN33)) & ((!(((((!(IN1)) & IN22) & (!(IN2))) & (!(IN3))) & IN21)) | IN14)) & ((!((((IN1 & IN22) & (!(IN2))) & (!(IN3))) & IN21)) | IN7)) & ((!(((((!(IN1)) & (!(IN22))) & IN2) & (!(IN3))) & IN21)) | IN32)) & ((!((((IN1 & (!(IN22))) & IN2) & (!(IN3))) & IN21)) | IN18)) & ((!(((((!(IN1)) & IN22) & IN2) & (!(IN3))) & IN21)) | IN30)) & ((!((((IN1 & IN22) & IN2) & (!(IN3))) & IN21)) | IN10)) & ((!(((((!(IN1)) & (!(IN22))) & (!(IN2))) & IN3) & IN21)) | IN17)) & ((!((((IN1 & (!(IN22))) & (!(IN2))) & IN3) & IN21)) | IN36)) & ((!(((((!(IN1)) & IN22) & (!(IN2))) & IN3) & IN21)) | IN16)) & ((!((((IN1 & IN22) & (!(IN2))) & IN3) & IN21)) | IN19)) & ((!(((((!(IN1)) & (!(IN22))) & IN2) & IN3) & IN21)) | IN12)) & ((!((((IN1 & (!(IN22))) & IN2) & IN3) & IN21)) | IN34)) & ((!(((((!(IN1)) & IN22) & IN2) & IN3) & IN21)) | IN37)) & ((!((((IN1 & IN22) & IN2) & IN3) & IN21)) | IN35)

*)

FUNCTION_BLOCK F_CollectInput
  VAR_IN_OUT
      Data : ARRAY[1..40] OF BOOL;
  END_VAR
  VAR_INPUT
      TICK  : BOOL := 0;
      IN1   : BOOL := 0;
      IN2   : BOOL := 0;
      IN3   : BOOL := 0;
      IN4   : BOOL := 0;
      IN5   : BOOL := 0;
      RESET : BOOL := FALSE;
  END_VAR
  VAR_OUTPUT
      Finished : BOOL;
  END_VAR
  VAR
      j    : USINT := 1;
      tock : BOOL  := 0;
  END_VAR
  IF NOT RESET AND tock = NOT TICK THEN
      Data[j]   := IN1;
      Data[j+1] := IN2;
      Data[j+2] := IN3;
      Data[j+3] := IN4;
      Data[j+4] := IN5;
      j := j + 5;
      tock := TICK;
  ELSE
      j := 1;
      tock := 0;
  END_IF;
  Finished := (j > 40);
END_FUNCTION_BLOCK

PROGRAM Boiler
  VAR
    Data  : ARRAY[1..40] OF BOOL;
    Ready : BOOL;
    CollectInput : F_CollectInput;
  END_VAR
  VAR
    TICK     AT %IX1.0 : BOOL;
    IN1      AT %IX0.3 : BOOL;
    IN2      AT %IX0.4 : BOOL;
    IN3      AT %IX0.5 : BOOL;
    IN4      AT %IX0.6 : BOOL;
    IN5      AT %IX0.7 : BOOL;
    OutReady AT %QX0.0 : BOOL := FALSE;
    FeedNext AT %QX0.1 : BOOL := FALSE;
    Out      AT %QX0.2 : BOOL;
  END_VAR
  CollectInput(TICK:=TICK, IN1:=IN1, IN2:=IN2, IN3:=IN3, IN4:=IN4, IN5:=IN5);
  Ready := CollectInput.Finished;
  FeedNext := 1;
  IF Ready THEN
    Out := (((((((((((((((((((((((((((((((((NOT (((((NOT Data[1]) AND (NOT Data[22])) AND (NOT Data[2])) AND (NOT Data[3])) AND (NOT Data[21]))) OR Data[23]) AND ((NOT ((((Data[1] AND (NOT Data[22])) AND (NOT Data[2])) AND (NOT Data[3])) AND (NOT Data[21]))) OR Data[5])) AND ((NOT (((((NOT Data[1]) AND Data[22]) AND (NOT Data[2])) AND (NOT Data[3])) AND (NOT Data[21]))) OR Data[4])) AND ((NOT ((((Data[1] AND Data[22]) AND (NOT Data[2])) AND (NOT Data[3])) AND (NOT Data[21]))) OR Data[6])) AND ((NOT (((((NOT Data[1]) AND (NOT Data[22])) AND Data[2]) AND (NOT Data[3])) AND (NOT Data[21]))) OR Data[8])) AND ((NOT ((((Data[1] AND (NOT Data[22])) AND Data[2]) AND (NOT Data[3])) AND (NOT Data[21]))) OR Data[20])) AND ((NOT (((((NOT Data[1]) AND Data[22]) AND Data[2]) AND (NOT Data[3])) AND (NOT Data[21]))) OR Data[24])) AND ((NOT ((((Data[1] AND Data[22]) AND Data[2]) AND (NOT Data[3])) AND (NOT Data[21]))) OR Data[26])) AND ((NOT (((((NOT Data[1]) AND (NOT Data[22])) AND (NOT Data[2])) AND Data[3]) AND (NOT Data[21]))) OR Data[25])) AND ((NOT ((((Data[1] AND (NOT Data[22])) AND (NOT Data[2])) AND Data[3]) AND (NOT Data[21]))) OR Data[27])) AND ((NOT (((((NOT Data[1]) AND Data[22]) AND (NOT Data[2])) AND Data[3]) AND (NOT Data[21]))) OR Data[13])) AND ((NOT ((((Data[1] AND Data[22]) AND (NOT Data[2])) AND Data[3]) AND (NOT Data[21]))) OR Data[11])) AND ((NOT (((((NOT Data[1]) AND (NOT Data[22])) AND Data[2]) AND Data[3]) AND (NOT Data[21]))) OR Data[9])) AND ((NOT ((((Data[1] AND (NOT Data[22])) AND Data[2]) AND Data[3]) AND (NOT Data[21]))) OR Data[15])) AND ((NOT (((((NOT Data[1]) AND Data[22]) AND Data[2]) AND Data[3]) AND (NOT Data[21]))) OR Data[31])) AND ((NOT ((((Data[1] AND Data[22]) AND Data[2]) AND Data[3]) AND (NOT Data[21]))) OR Data[28])) AND ((NOT (((((NOT Data[1]) AND (NOT Data[22])) AND (NOT Data[2])) AND (NOT Data[3])) AND Data[21])) OR Data[29])) AND ((NOT ((((Data[1] AND (NOT Data[22])) AND (NOT Data[2])) AND (NOT Data[3])) AND Data[21])) OR Data[33])) AND ((NOT (((((NOT Data[1]) AND Data[22]) AND (NOT Data[2])) AND (NOT Data[3])) AND Data[21])) OR Data[14])) AND ((NOT ((((Data[1] AND Data[22]) AND (NOT Data[2])) AND (NOT Data[3])) AND Data[21])) OR Data[7])) AND ((NOT (((((NOT Data[1]) AND (NOT Data[22])) AND Data[2]) AND (NOT Data[3])) AND Data[21])) OR Data[32])) AND ((NOT ((((Data[1] AND (NOT Data[22])) AND Data[2]) AND (NOT Data[3])) AND Data[21])) OR Data[18])) AND ((NOT (((((NOT Data[1]) AND Data[22]) AND Data[2]) AND (NOT Data[3])) AND Data[21])) OR Data[30])) AND ((NOT ((((Data[1] AND Data[22]) AND Data[2]) AND (NOT Data[3])) AND Data[21])) OR Data[10])) AND ((NOT (((((NOT Data[1]) AND (NOT Data[22])) AND (NOT Data[2])) AND Data[3]) AND Data[21])) OR Data[17])) AND ((NOT ((((Data[1] AND (NOT Data[22])) AND (NOT Data[2])) AND Data[3]) AND Data[21])) OR Data[36])) AND ((NOT (((((NOT Data[1]) AND Data[22]) AND (NOT Data[2])) AND Data[3]) AND Data[21])) OR Data[16])) AND ((NOT ((((Data[1] AND Data[22]) AND (NOT Data[2])) AND Data[3]) AND Data[21])) OR Data[19])) AND ((NOT (((((NOT Data[1]) AND (NOT Data[22])) AND Data[2]) AND Data[3]) AND Data[21])) OR Data[12])) AND ((NOT ((((Data[1] AND (NOT Data[22])) AND Data[2]) AND Data[3]) AND Data[21])) OR Data[34])) AND ((NOT (((((NOT Data[1]) AND Data[22]) AND Data[2]) AND Data[3]) AND Data[21])) OR Data[37])) AND ((NOT ((((Data[1] AND Data[22]) AND Data[2]) AND Data[3]) AND Data[21])) OR Data[35]));
    OutReady := 1;
    CollectInput(RESET:=TRUE);
  END_IF;
END_PROGRAM

CONFIGURATION Config0
  RESOURCE Res0 ON PLC
    TASK task0(INTERVAL := T#20ms,PRIORITY := 0);
    PROGRAM instance0 WITH task0 : Boiler;
  END_RESOURCE
END_CONFIGURATION

(* ---- 5-MUX_arity-tells-twixt.st ---- *)
(*
This code implements a shuffled multiplexer with 5 control bits.
The control bits are: Data[N3], Data[N1], Data[N5], Data[N20], Data[N22]
The input bits are: Data[N6], Data[N2], Data[N12], Data[N9], Data[N24], Data[N21], Data[N23], Data[N25], Data[N28], Data[N31], Data[N4], Data[N10], Data[N8], Data[N7], Data[N26], Data[N27], Data[N11], Data[N15], Data[N32], Data[N30], Data[N14], Data[N13], Data[N37], Data[N17], Data[N33], Data[N16], Data[N35], Data[N18], Data[N19], Data[N29], Data[N34], Data[N36]

The symbolic expression is:
((((((((((((((((((((((((((((((((!(((((!(IN3)) & (!(IN1))) & (!(IN5))) & (!(IN20))) & (!(IN22)))) | IN6) & ((!((((IN3 & (!(IN1))) & (!(IN5))) & (!(IN20))) & (!(IN22)))) | IN2)) & ((!(((((!(IN3)) & IN1) & (!(IN5))) & (!(IN20))) & (!(IN22)))) | IN12)) & ((!((((IN3 & IN1) & (!(IN5))) & (!(IN20))) & (!(IN22)))) | IN9)) & ((!(((((!(IN3)) & (!(IN1))) & IN5) & (!(IN20))) & (!(IN22)))) | IN24)) & ((!((((IN3 & (!(IN1))) & IN5) & (!(IN20))) & (!(IN22)))) | IN21)) & ((!(((((!(IN3)) & IN1) & IN5) & (!(IN20))) & (!(IN22)))) | IN23)) & ((!((((IN3 & IN1) & IN5) & (!(IN20))) & (!(IN22)))) | IN25)) & ((!(((((!(IN3)) & (!(IN1))) & (!(IN5))) & IN20) & (!(IN22)))) | IN28)) & ((!((((IN3 & (!(IN1))) & (!(IN5))) & IN20) & (!(IN22)))) | IN31)) & ((!(((((!(IN3)) & IN1) & (!(IN5))) & IN20) & (!(IN22)))) | IN4)) & ((!((((IN3 & IN1) & (!(IN5))) & IN20) & (!(IN22)))) | IN10)) & ((!(((((!(IN3)) & (!(IN1))) & IN5) & IN20) & (!(IN22)))) | IN8)) & ((!((((IN3 & (!(IN1))) & IN5) & IN20) & (!(IN22)))) | IN7)) & ((!(((((!(IN3)) & IN1) & IN5) & IN20) & (!(IN22)))) | IN26)) & ((!((((IN3 & IN1) & IN5) & IN20) & (!(IN22)))) | IN27)) & ((!(((((!(IN3)) & (!(IN1))) & (!(IN5))) & (!(IN20))) & IN22)) | IN11)) & ((!((((IN3 & (!(IN1))) & (!(IN5))) & (!(IN20))) & IN22)) | IN15)) & ((!(((((!(IN3)) & IN1) & (!(IN5))) & (!(IN20))) & IN22)) | IN32)) & ((!((((IN3 & IN1) & (!(IN5))) & (!(IN20))) & IN22)) | IN30)) & ((!(((((!(IN3)) & (!(IN1))) & IN5) & (!(IN20))) & IN22)) | IN14)) & ((!((((IN3 & (!(IN1))) & IN5) & (!(IN20))) & IN22)) | IN13)) & ((!(((((!(IN3)) & IN1) & IN5) & (!(IN20))) & IN22)) | IN37)) & ((!((((IN3 & IN1) & IN5) & (!(IN20))) & IN22)) | IN17)) & ((!(((((!(IN3)) & (!(IN1))) & (!(IN5))) & IN20) & IN22)) | IN33)) & ((!((((IN3 & (!(IN1))) & (!(IN5))) & IN20) & IN22)) | IN16)) & ((!(((((!(IN3)) & IN1) & (!(IN5))) & IN20) & IN22)) | IN35)) & ((!((((IN3 & IN1) & (!(IN5))) & IN20) & IN22)) | IN18)) & ((!(((((!(IN3)) & (!(IN1))) & IN5) & IN20) & IN22)) | IN19)) & ((!((((IN3 & (!(IN1))) & IN5) & IN20) & IN22)) | IN29)) & ((!(((((!(IN3)) & IN1) & IN5) & IN20) & IN22)) | IN34)) & ((!((((IN3 & IN1) & IN5) & IN20) & IN22)) | IN36)

*)

FUNCTION_BLOCK F_CollectInput
  VAR_IN_OUT
      Data : ARRAY[1..40] OF BOOL;
  END_VAR
  VAR_INPUT
      TICK  : BOOL := 0;
      IN1   : BOOL := 0;
      IN2   : BOOL := 0;
      IN3   : BOOL := 0;
      IN4   : BOOL := 0;
      IN5   : BOOL := 0;
      RESET : BOOL := FALSE;
  END_VAR
  VAR_OUTPUT
      Finished : BOOL;
  END_VAR
  VAR
      j    : USINT := 1;
      tock : BOOL  := 0;
  END_VAR
  IF NOT RESET AND tock = NOT TICK THEN
      Data[j]   := IN1;
      Data[j+1] := IN2;
      Data[j+2] := IN3;
      Data[j+3] := IN4;
      Data[j+4] := IN5;
      j := j + 5;
      tock := TICK;
  ELSE
      j := 1;
      tock := 0;
  END_IF;
  Finished := (j > 40);
END_FUNCTION_BLOCK

PROGRAM Boiler
  VAR
    Data  : ARRAY[1..40] OF BOOL;
    Ready : BOOL;
    CollectInput : F_CollectInput;
  END_VAR
  VAR
    TICK     AT %IX1.0 : BOOL;
    IN1      AT %IX0.3 : BOOL;
    IN2      AT %IX0.4 : BOOL;
    IN3      AT %IX0.5 : BOOL;
    IN4      AT %IX0.6 : BOOL;
    IN5      AT %IX0.7 : BOOL;
    OutReady AT %QX0.0 : BOOL := FALSE;
    FeedNext AT %QX0.1 : BOOL := FALSE;
    Out      AT %QX0.2 : BOOL;
  END_VAR
  CollectInput(TICK:=TICK, IN1:=IN1, IN2:=IN2, IN3:=IN3, IN4:=IN4, IN5:=IN5);
  Ready := CollectInput.Finished;
  FeedNext := 1;
  IF Ready THEN
    Out := (((((((((((((((((((((((((((((((((NOT (((((NOT Data[3]) AND (NOT Data[1])) AND (NOT Data[5])) AND (NOT Data[20])) AND (NOT Data[22]))) OR Data[6]) AND ((NOT ((((Data[3] AND (NOT Data[1])) AND (NOT Data[5])) AND (NOT Data[20])) AND (NOT Data[22]))) OR Data[2])) AND ((NOT (((((NOT Data[3]) AND Data[1]) AND (NOT Data[5])) AND (NOT Data[20])) AND (NOT Data[22]))) OR Data[12])) AND ((NOT ((((Data[3] AND Data[1]) AND (NOT Data[5])) AND (NOT Data[20])) AND (NOT Data[22]))) OR Data[9])) AND ((NOT (((((NOT Data[3]) AND (NOT Data[1])) AND Data[5]) AND (NOT Data[20])) AND (NOT Data[22]))) OR Data[24])) AND ((NOT ((((Data[3] AND (NOT Data[1])) AND Data[5]) AND (NOT Data[20])) AND (NOT Data[22]))) OR Data[21])) AND ((NOT (((((NOT Data[3]) AND Data[1]) AND Data[5]) AND (NOT Data[20])) AND (NOT Data[22]))) OR Data[23])) AND ((NOT ((((Data[3] AND Data[1]) AND Data[5]) AND (NOT Data[20])) AND (NOT Data[22]))) OR Data[25])) AND ((NOT (((((NOT Data[3]) AND (NOT Data[1])) AND (NOT Data[5])) AND Data[20]) AND (NOT Data[22]))) OR Data[28])) AND ((NOT ((((Data[3] AND (NOT Data[1])) AND (NOT Data[5])) AND Data[20]) AND (NOT Data[22]))) OR Data[31])) AND ((NOT (((((NOT Data[3]) AND Data[1]) AND (NOT Data[5])) AND Data[20]) AND (NOT Data[22]))) OR Data[4])) AND ((NOT ((((Data[3] AND Data[1]) AND (NOT Data[5])) AND Data[20]) AND (NOT Data[22]))) OR Data[10])) AND ((NOT (((((NOT Data[3]) AND (NOT Data[1])) AND Data[5]) AND Data[20]) AND (NOT Data[22]))) OR Data[8])) AND ((NOT ((((Data[3] AND (NOT Data[1])) AND Data[5]) AND Data[20]) AND (NOT Data[22]))) OR Data[7])) AND ((NOT (((((NOT Data[3]) AND Data[1]) AND Data[5]) AND Data[20]) AND (NOT Data[22]))) OR Data[26])) AND ((NOT ((((Data[3] AND Data[1]) AND Data[5]) AND Data[20]) AND (NOT Data[22]))) OR Data[27])) AND ((NOT (((((NOT Data[3]) AND (NOT Data[1])) AND (NOT Data[5])) AND (NOT Data[20])) AND Data[22])) OR Data[11])) AND ((NOT ((((Data[3] AND (NOT Data[1])) AND (NOT Data[5])) AND (NOT Data[20])) AND Data[22])) OR Data[15])) AND ((NOT (((((NOT Data[3]) AND Data[1]) AND (NOT Data[5])) AND (NOT Data[20])) AND Data[22])) OR Data[32])) AND ((NOT ((((Data[3] AND Data[1]) AND (NOT Data[5])) AND (NOT Data[20])) AND Data[22])) OR Data[30])) AND ((NOT (((((NOT Data[3]) AND (NOT Data[1])) AND Data[5]) AND (NOT Data[20])) AND Data[22])) OR Data[14])) AND ((NOT ((((Data[3] AND (NOT Data[1])) AND Data[5]) AND (NOT Data[20])) AND Data[22])) OR Data[13])) AND ((NOT (((((NOT Data[3]) AND Data[1]) AND Data[5]) AND (NOT Data[20])) AND Data[22])) OR Data[37])) AND ((NOT ((((Data[3] AND Data[1]) AND Data[5]) AND (NOT Data[20])) AND Data[22])) OR Data[17])) AND ((NOT (((((NOT Data[3]) AND (NOT Data[1])) AND (NOT Data[5])) AND Data[20]) AND Data[22])) OR Data[33])) AND ((NOT ((((Data[3] AND (NOT Data[1])) AND (NOT Data[5])) AND Data[20]) AND Data[22])) OR Data[16])) AND ((NOT (((((NOT Data[3]) AND Data[1]) AND (NOT Data[5])) AND Data[20]) AND Data[22])) OR Data[35])) AND ((NOT ((((Data[3] AND Data[1]) AND (NOT Data[5])) AND Data[20]) AND Data[22])) OR Data[18])) AND ((NOT (((((NOT Data[3]) AND (NOT Data[1])) AND Data[5]) AND Data[20]) AND Data[22])) OR Data[19])) AND ((NOT ((((Data[3] AND (NOT Data[1])) AND Data[5]) AND Data[20]) AND Data[22])) OR Data[29])) AND ((NOT (((((NOT Data[3]) AND Data[1]) AND Data[5]) AND Data[20]) AND Data[22])) OR Data[34])) AND ((NOT ((((Data[3] AND Data[1]) AND Data[5]) AND Data[20]) AND Data[22])) OR Data[36]));
    OutReady := 1;
    CollectInput(RESET:=TRUE);
  END_IF;
END_PROGRAM

CONFIGURATION Config0
  RESOURCE Res0 ON PLC
    TASK task0(INTERVAL := T#20ms,PRIORITY := 0);
    PROGRAM instance0 WITH task0 : Boiler;
  END_RESOURCE
END_CONFIGURATION
